// TwinCAT 3 PLC project KFEArbiter
// Title: KFE-ARBITER
// Company: SLAC - LCLS
// ProjectVersion: 0.0.0
// ProgramVersion: 3.1.4022.7
// CompilerDefines: K
// libraries:
//   PMPS, * (SLAC - LCLS)
//   Tc2_Math, * (Beckhoff Automation GmbH)
//   Tc2_MC2, * (Beckhoff Automation GmbH)
//   Tc2_Standard, * (Beckhoff Automation GmbH)
//   Tc2_System, * (Beckhoff Automation GmbH)
//   Tc2_SystemCX, * (Beckhoff Automation GmbH)
//   Tc2_Utilities, * (Beckhoff Automation GmbH)
//   Tc3_Module, * (Beckhoff Automation GmbH)
//   LCLS General,2.8.2,SLAC
// project tree:
//   / FFOTask.TcTTO, PlcTask.TcTTO
//   GVLs/ GVL.TcGVL, GVL_CheckBounds.TcGVL
//   ImplicitChecks/ CheckBounds.TcPOU, CheckRangeSigned.TcPOU, CheckRangeUnsigned.TcPOU
//   POUs/ CurrentBPUpdate.TcPOU, CXDisplay.TcPOU, Fast_Faults_Evaluate.TcPOU, FB_BeamClassOutputs.TcPOU, MachineSimulation.TcPOU, MAIN.TcPOU, PMPS_Arbiter.TcPOU, P_AT1K0_SL1K0.TcPOU, P_BeamClassAssertion.TcPOU, P_Override_Tran_BC.TcPOU, P_SATT.TcPOU, Testing.TcPOU
//   POUs/TEMP/ FB_ArbiterToSubSys_IO.TcPOU
// real-time tasks:
//   TASK PlcTask: cycle T#10ms, priority 2, ADS port 350
//   TASK FFOTask: cycle T#1ms, priority 1, ADS port 351
// I/O:
//   DEVICE Device 1 (EtherCAT), AmsNetId 0.0.0.0.2.1
//     E0 (EK1200) [EK1200-5000 EtherCAT Power supply (2A E-Bus)]
//       FFO [EL2202 2Ch. Dig. Output 24V, 0.5A]
//       PMPS_Premp [EL2809 16Ch. Dig. Output 24V, 0.5A]
//       E3 (EK1122) [EK1122 2 port EtherCAT junction]
//         950-101W-R4-MPS-2 [EK1100 EtherCAT Coupler (2A E-Bus)]
//           PPS Stoppers 1 [EL1008 8Ch. Dig. Input 24V, 3ms]
//           PPS Stoppers 2 [EL1008 8Ch. Dig. Input 24V, 3ms]
//           950-101W-R4-MPS-2-E3 (EL9011) [EL9011 End Terminal]
//       Term 22 (EK1110) [EK1110 EtherCAT extension]
//     B940-009-R07-MPS-1 CU1-ESC1 [CU1128 6x EtherCAT junction]
//       plc-kfe-motion [EL6695 EtherCAT Bridge terminal (Secondary)]
//       plc-kfe-gmd-vac-01 [EL6695 EtherCAT Bridge terminal (Secondary)]
//       plc-kfe-xgmd-vac-01 [EL6695 EtherCAT Bridge terminal (Secondary)]
//       plc-kfe-vac [EL6692 EtherCAT Bridge terminal (Secondary)]
//       plc-kfe-gatt [EL6695 EtherCAT Bridge terminal (Secondary)]
//       plc-tmo-mot [EL6692 EtherCAT Bridge terminal (Secondary)]
//       plc-tmo-optics [EL6695 EtherCAT Bridge terminal (Secondary)]
//       plc-tmo-vac [EL6692 EtherCAT Bridge terminal (Secondary)]
//       B940-009-R07-MPS-1 CU1-ESC2 [CU1128 6x EtherCAT junction - Dev A]
//         plc-rix-mot
//         plc-rix-vac
//         plc-rix-optics
//         plc-crix-vac
//         plc-crix-mot
//       B940-009-R07-MPS-1 CU1-ESC3 [CU1128 6x EtherCAT junction - Dev B]
//         plc-qrix-vac
//         plc-qrix-mot
//         plc-txi-optics
//     plc-txi-mot [EL6695 EtherCAT Bridge terminal (Secondary)]
//     plc-txi-vac [EL6695 EtherCAT Bridge terminal (Secondary)]
// variable links:
//   KFEArbiter Instance <-> Device 1 (EtherCAT)
//     PlcTask Inputs/MAIN.fbEcatDiag.arrEcMasterNetId <-> InfoData/AmsNetId
//     PlcTask Inputs/MAIN.fbEcatDiag.nEcMasterDevState <-> Inputs/DevState
//     PlcTask Inputs/MAIN.fbEcatDiag.nEcMasterDeviceId <-> InfoData/DevId
//     PlcTask Inputs/MAIN.fbEcatDiag.nEcMasterSlaveCount <-> Inputs/SlaveCount
//     PlcTask Inputs/MAIN.fbEcatDiag.nEcMasterSlaveCountCfg <-> InfoData/CfgSlaveCount
//     PlcTask Inputs/MAIN.fbEcatDiag.wFrmXWcState <-> Inputs/Frm1WcState
//   KFEArbiter Instance <-> Device 1 (EtherCAT)/B940-009-R07-MPS-1 CU1-ESC1/B940-009-R07-MPS-1 CU1-ESC2/plc-crix-mot
//     PlcTask Inputs/PMPS_Arbiter.plc_crix_mot_PMPS_IO.i_Connected <-> SYNC Inputs/External device not connected
//     PlcTask Inputs/PMPS_Arbiter.plc_crix_mot_PMPS_IO.i_RequestedBP <-> IO Inputs/RequestedBP
//     PlcTask Inputs/PMPS_Arbiter.plc_crix_mot_PMPS_IO.i_TxPDOState <-> SYNC Inputs/TxPDO state
//     PlcTask Inputs/PMPS_Arbiter.plc_crix_mot_PMPS_IO.i_WcState <-> WcState/WcStateIn
//     PlcTask Outputs/PMPS_Arbiter.plc_crix_mot_PMPS_IO.o_CurrentBP <-> IO Outputs/CurrentBP
//   KFEArbiter Instance <-> Device 1 (EtherCAT)/B940-009-R07-MPS-1 CU1-ESC1/B940-009-R07-MPS-1 CU1-ESC2/plc-crix-vac
//     PlcTask Inputs/PMPS_Arbiter.plc_crix_vac_PMPS_IO.i_Connected <-> SYNC Inputs/External device not connected
//     PlcTask Inputs/PMPS_Arbiter.plc_crix_vac_PMPS_IO.i_RequestedBP <-> IO Inputs/RequestedBP
//     PlcTask Inputs/PMPS_Arbiter.plc_crix_vac_PMPS_IO.i_TxPDOState <-> SYNC Inputs/TxPDO state
//     PlcTask Inputs/PMPS_Arbiter.plc_crix_vac_PMPS_IO.i_WcState <-> WcState/WcStateIn
//     PlcTask Outputs/PMPS_Arbiter.plc_crix_vac_PMPS_IO.o_CurrentBP <-> IO Outputs/CurrentBP
//   KFEArbiter Instance <-> Device 1 (EtherCAT)/B940-009-R07-MPS-1 CU1-ESC1/B940-009-R07-MPS-1 CU1-ESC2/plc-rix-mot
//     PlcTask Inputs/PMPS_Arbiter.plc_rix_mot_PMPS_IO.i_Connected <-> SYNC Inputs/External device not connected
//     PlcTask Inputs/PMPS_Arbiter.plc_rix_mot_PMPS_IO.i_RequestedBP <-> IO Inputs/RequestedBP
//     PlcTask Inputs/PMPS_Arbiter.plc_rix_mot_PMPS_IO.i_TxPDOState <-> SYNC Inputs/TxPDO state
//     PlcTask Inputs/PMPS_Arbiter.plc_rix_mot_PMPS_IO.i_WcState <-> WcState/WcStateIn
//     PlcTask Inputs/P_SATT.i_SattArrayStatus_RIX <-> IO Inputs/SattArrayStatus
//     PlcTask Inputs/P_SATT.i_bWcStateIn_rix_mot <-> WcState/WcStateIn
//     PlcTask Inputs/P_SATT.i_bWcStateOut_rix_mot <-> WcState/WcStateOut
//     PlcTask Inputs/P_SATT.i_nState_rix_mot <-> InfoData/State
//     PlcTask Outputs/PMPS_Arbiter.plc_rix_mot_PMPS_IO.o_CurrentBP <-> IO Outputs/CurrentBP
//     PlcTask Outputs/P_SATT.q_SattArrayReq <-> IO Outputs/SattArrayReq
//   KFEArbiter Instance <-> Device 1 (EtherCAT)/B940-009-R07-MPS-1 CU1-ESC1/B940-009-R07-MPS-1 CU1-ESC2/plc-rix-optics
//     PlcTask Inputs/CurrentBPUpdate.i_MR1K1_ENC <-> IO Inputs/MR1K1_Y_ENC
//     PlcTask Inputs/PMPS_Arbiter.plc_rix_optics_PMPS_IO.i_Connected <-> SYNC Inputs/External device not connected
//     PlcTask Inputs/PMPS_Arbiter.plc_rix_optics_PMPS_IO.i_RequestedBP <-> IO Inputs/RequestedBP
//     PlcTask Inputs/PMPS_Arbiter.plc_rix_optics_PMPS_IO.i_TxPDOState <-> SYNC Inputs/TxPDO state
//     PlcTask Inputs/PMPS_Arbiter.plc_rix_optics_PMPS_IO.i_WcState <-> WcState/WcStateIn
//     PlcTask Outputs/PMPS_Arbiter.plc_rix_optics_PMPS_IO.o_CurrentBP <-> IO Outputs/CurrentBP
//   KFEArbiter Instance <-> Device 1 (EtherCAT)/B940-009-R07-MPS-1 CU1-ESC1/B940-009-R07-MPS-1 CU1-ESC2/plc-rix-vac
//     PlcTask Inputs/PMPS_Arbiter.plc_rix_vac_PMPS_IO.i_Connected <-> SYNC Inputs/External device not connected
//     PlcTask Inputs/PMPS_Arbiter.plc_rix_vac_PMPS_IO.i_RequestedBP <-> IO Inputs/RequestedBP
//     PlcTask Inputs/PMPS_Arbiter.plc_rix_vac_PMPS_IO.i_TxPDOState <-> SYNC Inputs/TxPDO state
//     PlcTask Inputs/PMPS_Arbiter.plc_rix_vac_PMPS_IO.i_WcState <-> WcState/WcStateIn
//     PlcTask Outputs/PMPS_Arbiter.plc_rix_vac_PMPS_IO.o_CurrentBP <-> IO Outputs/CurrentBP
//   KFEArbiter Instance <-> Device 1 (EtherCAT)/B940-009-R07-MPS-1 CU1-ESC1/B940-009-R07-MPS-1 CU1-ESC3/plc-qrix-mot
//     PlcTask Inputs/PMPS_Arbiter.plc_qrix_mot_PMPS_IO.i_Connected <-> SYNC Inputs/External device not connected
//     PlcTask Inputs/PMPS_Arbiter.plc_qrix_mot_PMPS_IO.i_RequestedBP <-> IO Inputs/RequestedBP
//     PlcTask Inputs/PMPS_Arbiter.plc_qrix_mot_PMPS_IO.i_TxPDOState <-> SYNC Inputs/TxPDO state
//     PlcTask Inputs/PMPS_Arbiter.plc_qrix_mot_PMPS_IO.i_WcState <-> WcState/WcStateIn
//     PlcTask Outputs/PMPS_Arbiter.plc_qrix_mot_PMPS_IO.o_CurrentBP <-> IO Outputs/CurrentBP
//   KFEArbiter Instance <-> Device 1 (EtherCAT)/B940-009-R07-MPS-1 CU1-ESC1/B940-009-R07-MPS-1 CU1-ESC3/plc-qrix-vac
//     PlcTask Inputs/Fast_Faults_Evaluate.i_xFastFaultOut_qrix_vac <-> IO Inputs/FFO
//     PlcTask Inputs/PMPS_Arbiter.plc_qrix_vac_PMPS_IO.i_Connected <-> SYNC Inputs/External device not connected
//     PlcTask Inputs/PMPS_Arbiter.plc_qrix_vac_PMPS_IO.i_RequestedBP <-> IO Inputs/RequestedBP
//     PlcTask Inputs/PMPS_Arbiter.plc_qrix_vac_PMPS_IO.i_TxPDOState <-> SYNC Inputs/TxPDO state
//     PlcTask Inputs/PMPS_Arbiter.plc_qrix_vac_PMPS_IO.i_WcState <-> WcState/WcStateIn
//     PlcTask Outputs/PMPS_Arbiter.plc_qrix_vac_PMPS_IO.o_CurrentBP <-> IO Outputs/CurrentBP
//   KFEArbiter Instance <-> Device 1 (EtherCAT)/B940-009-R07-MPS-1 CU1-ESC1/B940-009-R07-MPS-1 CU1-ESC3/plc-txi-optics
//     PlcTask Inputs/CurrentBPUpdate.i_MR1K3_ENC <-> IO Inputs/MR1K3_Y_ENC
//     PlcTask Inputs/CurrentBPUpdate.i_MR2K3_ENC <-> IO Inputs/MR2K3_Y_ENC
//     PlcTask Inputs/Fast_Faults_Evaluate.i_xFastFaultOut_txi_optics <-> IO Inputs/FFO
//     PlcTask Inputs/PMPS_Arbiter.plc_txi_optics_PMPS_IO.i_Connected <-> SYNC Inputs/External device not connected
//     PlcTask Inputs/PMPS_Arbiter.plc_txi_optics_PMPS_IO.i_RequestedBP <-> IO Inputs/RequestedBP
//     PlcTask Inputs/PMPS_Arbiter.plc_txi_optics_PMPS_IO.i_TxPDOState <-> SYNC Inputs/TxPDO state
//     PlcTask Inputs/PMPS_Arbiter.plc_txi_optics_PMPS_IO.i_WcState <-> WcState/WcStateIn
//     PlcTask Outputs/PMPS_Arbiter.plc_txi_optics_PMPS_IO.o_CurrentBP <-> IO Outputs/CurrentBP
//   KFEArbiter Instance <-> Device 1 (EtherCAT)/B940-009-R07-MPS-1 CU1-ESC1/plc-kfe-gatt
//     PlcTask Inputs/PMPS_Arbiter.plc_kfe_gatt_PMPS_IO.i_Connected <-> SYNC Inputs/External device not connected
//     PlcTask Inputs/PMPS_Arbiter.plc_kfe_gatt_PMPS_IO.i_RequestedBP <-> IO Inputs/RequestedBP
//     PlcTask Inputs/PMPS_Arbiter.plc_kfe_gatt_PMPS_IO.i_TxPDOState <-> SYNC Inputs/TxPDO state
//     PlcTask Inputs/PMPS_Arbiter.plc_kfe_gatt_PMPS_IO.i_WcState <-> WcState/WcStateIn
//     PlcTask Inputs/P_AT1K0_SL1K0.i_bWcStateIn_AT1K0 <-> WcState/WcStateIn
//     PlcTask Inputs/P_AT1K0_SL1K0.i_bWcStateOut_AT1K0 <-> WcState/WcStateOut
//     PlcTask Inputs/P_AT1K0_SL1K0.i_nState_AT1K0 <-> InfoData/State
//     PlcTask Inputs/P_AT1K0_SL1K0.i_nTranToAT1K0Stat <-> IO Inputs/Current Transmission
//     PlcTask Outputs/PMPS_Arbiter.plc_kfe_gatt_PMPS_IO.o_CurrentBP <-> IO Outputs/CurrentBP
//     PlcTask Outputs/P_AT1K0_SL1K0.q_nTranToAT1K0Req <-> IO Outputs/Requested Transmission
//   KFEArbiter Instance <-> Device 1 (EtherCAT)/B940-009-R07-MPS-1 CU1-ESC1/plc-kfe-gmd-vac-01
//     PlcTask Inputs/PMPS_Arbiter.plc_kfe_gmd_PMPS_IO.i_Connected <-> SYNC Inputs/External device not connected
//     PlcTask Inputs/PMPS_Arbiter.plc_kfe_gmd_PMPS_IO.i_RequestedBP <-> IO Inputs/RequestedBP
//     PlcTask Inputs/PMPS_Arbiter.plc_kfe_gmd_PMPS_IO.i_TxPDOState <-> SYNC Inputs/TxPDO state
//     PlcTask Inputs/PMPS_Arbiter.plc_kfe_gmd_PMPS_IO.i_WcState <-> WcState/WcStateIn
//     PlcTask Outputs/PMPS_Arbiter.plc_kfe_gmd_PMPS_IO.o_CurrentBP <-> IO Outputs/CurrentBP
//   KFEArbiter Instance <-> Device 1 (EtherCAT)/B940-009-R07-MPS-1 CU1-ESC1/plc-kfe-motion
//     PlcTask Inputs/CurrentBPUpdate.ST1K4_Y_ENC <-> IO Inputs/ST1K4_Y_ENC
//     PlcTask Inputs/PMPS_Arbiter.plc_kfe_motion_PMPS_IO.i_Connected <-> SYNC Inputs/External device not connected
//     PlcTask Inputs/PMPS_Arbiter.plc_kfe_motion_PMPS_IO.i_RequestedBP <-> IO Inputs/RequestedBP
//     PlcTask Inputs/PMPS_Arbiter.plc_kfe_motion_PMPS_IO.i_TxPDOState <-> SYNC Inputs/TxPDO state
//     PlcTask Inputs/PMPS_Arbiter.plc_kfe_motion_PMPS_IO.i_WcState <-> WcState/WcStateIn
//     PlcTask Inputs/P_AT1K0_SL1K0.i_bWcStateIn_KFEMOT <-> WcState/WcStateIn
//     PlcTask Inputs/P_AT1K0_SL1K0.i_bWcStateOut_KFEMOT <-> WcState/WcStateOut
//     PlcTask Inputs/P_AT1K0_SL1K0.i_nState_KFEMOT <-> InfoData/State
//     PlcTask Inputs/P_AT1K0_SL1K0.i_stAptArrayStat <-> IO Inputs/AptArrayStatus
//     PlcTask Inputs/P_SATT.i_SattArrayStatus_KFE <-> IO Inputs/SattArrayStatus
//     PlcTask Inputs/P_SATT.i_bWcStateIn_kfe_mot <-> WcState/WcStateIn
//     PlcTask Inputs/P_SATT.i_bWcStateOut_kfe_mot <-> WcState/WcStateOut
//     PlcTask Inputs/P_SATT.i_nState_kfe_mot <-> InfoData/State
//     PlcTask Outputs/PMPS_Arbiter.plc_kfe_motion_PMPS_IO.o_CurrentBP <-> IO Outputs/CurrentBP
//     PlcTask Outputs/P_AT1K0_SL1K0.q_stAptArrayReq <-> IO Outputs/AptArrayReq
//   KFEArbiter Instance <-> Device 1 (EtherCAT)/B940-009-R07-MPS-1 CU1-ESC1/plc-kfe-vac
//     PlcTask Inputs/PMPS_Arbiter.plc_kfe_vac_PMPS_IO.i_Connected <-> SYNC Inputs/External device not connected
//     PlcTask Inputs/PMPS_Arbiter.plc_kfe_vac_PMPS_IO.i_RequestedBP <-> IO Inputs/RequestedBP
//     PlcTask Inputs/PMPS_Arbiter.plc_kfe_vac_PMPS_IO.i_TxPDOState <-> SYNC Inputs/TxPDO state
//     PlcTask Inputs/PMPS_Arbiter.plc_kfe_vac_PMPS_IO.i_WcState <-> WcState/WcStateIn
//     PlcTask Outputs/PMPS_Arbiter.plc_kfe_vac_PMPS_IO.o_CurrentBP <-> IO Outputs/CurrentBP
//   KFEArbiter Instance <-> Device 1 (EtherCAT)/B940-009-R07-MPS-1 CU1-ESC1/plc-kfe-xgmd-vac-01
//     PlcTask Inputs/PMPS_Arbiter.plc_kfe_xgmd_PMPS_IO.i_Connected <-> SYNC Inputs/External device not connected
//     PlcTask Inputs/PMPS_Arbiter.plc_kfe_xgmd_PMPS_IO.i_RequestedBP <-> IO Inputs/RequestedBP
//     PlcTask Inputs/PMPS_Arbiter.plc_kfe_xgmd_PMPS_IO.i_TxPDOState <-> SYNC Inputs/TxPDO state
//     PlcTask Inputs/PMPS_Arbiter.plc_kfe_xgmd_PMPS_IO.i_WcState <-> WcState/WcStateIn
//     PlcTask Outputs/PMPS_Arbiter.plc_kfe_xgmd_PMPS_IO.o_CurrentBP <-> IO Outputs/CurrentBP
//   KFEArbiter Instance <-> Device 1 (EtherCAT)/B940-009-R07-MPS-1 CU1-ESC1/plc-tmo-mot
//     PlcTask Inputs/CurrentBPUpdate.st4k4Watcher.i_StopperInLS <-> IO Inputs/bST4K4_IN
//     PlcTask Inputs/CurrentBPUpdate.st4k4Watcher.i_StopperOutLS <-> IO Inputs/bST4K4_OUT
//     PlcTask Inputs/PMPS_Arbiter.plc_tmo_motion_PMPS_IO.i_Connected <-> SYNC Inputs/External device not connected
//     PlcTask Inputs/PMPS_Arbiter.plc_tmo_motion_PMPS_IO.i_RequestedBP <-> IO Inputs/RequestedBP
//     PlcTask Inputs/PMPS_Arbiter.plc_tmo_motion_PMPS_IO.i_TxPDOState <-> SYNC Inputs/TxPDO state
//     PlcTask Inputs/PMPS_Arbiter.plc_tmo_motion_PMPS_IO.i_WcState <-> WcState/WcStateIn
//     PlcTask Outputs/PMPS_Arbiter.plc_tmo_motion_PMPS_IO.o_CurrentBP <-> IO Outputs/CurrentBP
//   KFEArbiter Instance <-> Device 1 (EtherCAT)/B940-009-R07-MPS-1 CU1-ESC1/plc-tmo-optics
//     PlcTask Inputs/PMPS_Arbiter.plc_tmo_optics_PMPS_IO.i_Connected <-> SYNC Inputs/External device not connected
//     PlcTask Inputs/PMPS_Arbiter.plc_tmo_optics_PMPS_IO.i_RequestedBP <-> IO Inputs/RequestedBP
//     PlcTask Inputs/PMPS_Arbiter.plc_tmo_optics_PMPS_IO.i_TxPDOState <-> SYNC Inputs/TxPDO state
//     PlcTask Inputs/PMPS_Arbiter.plc_tmo_optics_PMPS_IO.i_WcState <-> WcState/WcStateIn
//     PlcTask Outputs/PMPS_Arbiter.plc_tmo_optics_PMPS_IO.o_CurrentBP <-> IO Outputs/CurrentBP
//   KFEArbiter Instance <-> Device 1 (EtherCAT)/B940-009-R07-MPS-1 CU1-ESC1/plc-tmo-vac
//     PlcTask Inputs/PMPS_Arbiter.plc_tmo_vacuum_PMPS_IO.i_Connected <-> SYNC Inputs/External device not connected
//     PlcTask Inputs/PMPS_Arbiter.plc_tmo_vacuum_PMPS_IO.i_RequestedBP <-> IO Inputs/RequestedBP
//     PlcTask Inputs/PMPS_Arbiter.plc_tmo_vacuum_PMPS_IO.i_TxPDOState <-> SYNC Inputs/TxPDO state
//     PlcTask Inputs/PMPS_Arbiter.plc_tmo_vacuum_PMPS_IO.i_WcState <-> WcState/WcStateIn
//     PlcTask Outputs/PMPS_Arbiter.plc_tmo_vacuum_PMPS_IO.o_CurrentBP <-> IO Outputs/CurrentBP
//   KFEArbiter Instance <-> Device 1 (EtherCAT)/E0 (EK1200)/E3 (EK1122)/950-101W-R4-MPS-2/PPS Stoppers 1
//     PlcTask Inputs/CurrentBPUpdate.st1k2Watcher.i_StopperInLS <-> Channel 3/ST1K2 IN
//     PlcTask Inputs/CurrentBPUpdate.st1k3Watcher.i_StopperInLS <-> Channel 5/ST1K3 IN
//     PlcTask Inputs/CurrentBPUpdate.st3k4Watcher.i_StopperInLS <-> Channel 1/ST3K4 IN
//     PlcTask Inputs/CurrentBPUpdate.st1k2Watcher.i_StopperOutLS <-> Channel 4/ST1K2 OUT
//     PlcTask Inputs/CurrentBPUpdate.st1k3Watcher.i_StopperOutLS <-> Channel 6/ST1K3 OUT
//     PlcTask Inputs/CurrentBPUpdate.st3k4Watcher.i_StopperOutLS <-> Channel 2/ST3K4 OUT
//   KFEArbiter Instance <-> Device 1 (EtherCAT)/E0 (EK1200)/FFO
//     PlcTask Outputs/GVL.g_FastFaultOutput1.q_xFastFaultOut <-> Channel 1/Output
//     PlcTask Outputs/GVL.g_FastFaultOutput2.q_xFastFaultOut <-> Channel 2/Output
//   KFEArbiter Instance <-> Device 1 (EtherCAT)/E0 (EK1200)/PMPS_Premp
//     PlcTask Outputs/CurrentBPUpdate.q_MR1K1_VETO <-> Channel 13/MR1K1 IN
//     PlcTask Outputs/CurrentBPUpdate.st1k2Watcher.q_StopperIN_Relay <-> Channel 14/ST1K2 RELAY IN
//     PlcTask Outputs/CurrentBPUpdate.st1k3Watcher.q_StopperIN_Relay <-> Channel 7/ST1K3 RELAY IN
//     PlcTask Outputs/CurrentBPUpdate.st3k4Watcher.q_StopperIN_Relay <-> Channel 12/ST3K4 RELAY IN
//     PlcTask Outputs/MAIN.bM1K1_OUT_Override <-> Channel 8/Output
//     PlcTask Outputs/PMPS_Arbiter.fbCuInterface.q_CLTS_ASSERTION_LINES[1] <-> Channel 9/Output
//     PlcTask Outputs/PMPS_Arbiter.fbCuInterface.q_CLTS_ASSERTION_LINES[2] <-> Channel 10/Output
//     PlcTask Outputs/PMPS_Arbiter.fbCuInterface.q_CLTS_ASSERTION_LINES[3] <-> Channel 11/Output
//     PlcTask Outputs/P_BeamClassAssertion.fbMPSInterface.q_BC_ASSERTION_LINES[{1..4}] <-> Channel {1..4}/Output  (4 links)
//   KFEArbiter Instance <-> Device 1 (EtherCAT)/plc-txi-mot
//     PlcTask Inputs/Fast_Faults_Evaluate.i_xFastFaultOut_txi_mot <-> IO Inputs/FFO
//     PlcTask Inputs/PMPS_Arbiter.plc_txi_motion_PMPS_IO.i_Connected <-> SYNC Inputs/External device not connected
//     PlcTask Inputs/PMPS_Arbiter.plc_txi_motion_PMPS_IO.i_RequestedBP <-> IO Inputs/RequestedBP
//     PlcTask Inputs/PMPS_Arbiter.plc_txi_motion_PMPS_IO.i_TxPDOState <-> SYNC Inputs/TxPDO state
//     PlcTask Inputs/PMPS_Arbiter.plc_txi_motion_PMPS_IO.i_WcState <-> WcState/WcStateIn
//     PlcTask Outputs/PMPS_Arbiter.plc_txi_motion_PMPS_IO.o_CurrentBP <-> IO Outputs/CurrentBP
//   KFEArbiter Instance <-> Device 1 (EtherCAT)/plc-txi-vac
//     PlcTask Inputs/Fast_Faults_Evaluate.i_xFastFaultOut_txi_vac <-> IO Inputs/FFO
//     PlcTask Inputs/PMPS_Arbiter.plc_txi_vacuum_PMPS_IO.i_Connected <-> SYNC Inputs/External device not connected
//     PlcTask Inputs/PMPS_Arbiter.plc_txi_vacuum_PMPS_IO.i_RequestedBP <-> IO Inputs/RequestedBP
//     PlcTask Inputs/PMPS_Arbiter.plc_txi_vacuum_PMPS_IO.i_TxPDOState <-> SYNC Inputs/TxPDO state
//     PlcTask Inputs/PMPS_Arbiter.plc_txi_vacuum_PMPS_IO.i_WcState <-> WcState/WcStateIn
//     PlcTask Outputs/PMPS_Arbiter.plc_txi_vacuum_PMPS_IO.o_CurrentBP <-> IO Outputs/CurrentBP

CONFIGURATION KFEArbiter
    RESOURCE PLC ON TwinCAT3
        TASK FFOTask(INTERVAL := T#1ms, PRIORITY := 1);
        TASK PlcTask(INTERVAL := T#10ms, PRIORITY := 2);
        PROGRAM MAIN WITH PlcTask : MAIN;
    END_RESOURCE
END_CONFIGURATION

// ---- GVLs/GVL.TcGVL

VAR_GLOBAL
   {attribute 'pytmc' := '
    pv: @(PREFIX)Arbiter:01
    '}
    g_fbArbiter1	:	FB_Arbiter(25);

    {attribute 'pytmc' := '
    pv: @(PREFIX)Arbiter:02
    '}
    g_fbArbiter2	:	FB_Arbiter(25); //Used to line beam parameter

    ReqBP	:	ST_BeamParams; //Currently the placeholder for the fully arbitrated BP set

    // These are added for the additional low selector to figure out the override
    stArbiter1BP:ST_BeamParams; // a place holder for the arbitrated safe beam set from all the connected PLCs
    stCurrentFakeBP:ST_BeamParams; //Currently the placeholder for the fake arbitrated BP set to go to the rest of the PLC

    {attribute 'pytmc' := '
    pv: @(PREFIX)FFO:01
    '}
    {attribute 'TcLinkTo' := '.q_xFastFaultOut:=TIIB[FFO]^Channel 1^Output'}
    g_FastFaultOutput1	:	FB_HardwareFFOutput := (bAutoReset:=TRUE);

    {attribute 'pytmc' := '
    pv: @(PREFIX)FFO:02
    '}
    {attribute 'TcLinkTo' := '.q_xFastFaultOut:=TIIB[FFO]^Channel 2^Output'}
    g_FastFaultOutput2	:	FB_HardwareFFOutput := (bAutoReset:=TRUE);
	
	
	//The following faults will be per hutch and vetoed by the hutch specific veto
	//TMO OPTICS, VAC and Motion, DREAM
	{attribute 'pytmc' := '
    pv: @(PREFIX)FFO:03
    '}
    g_FastFaultOutput3	:	FB_HardwareFFOutput := (bAutoReset:=TRUE);
	{attribute 'pytmc' := '
    pv: @(PREFIX)FFO:04
    '}
    g_FastFaultOutput4	:	FB_HardwareFFOutput := (bAutoReset:=TRUE);
	
	
	//RIX Motion, QRIX and CRIX
	//NOTE: NOT OPTICS, NO VETO for OPTICS
	{attribute 'pytmc' := '
    pv: @(PREFIX)FFO:05
    '}
    g_FastFaultOutput5	:	FB_HardwareFFOutput := (bAutoReset:=TRUE);
	
	{attribute 'pytmc' := '
    pv: @(PREFIX)FFO:06
    '}
    g_FastFaultOutput6	:	FB_HardwareFFOutput := (bAutoReset:=TRUE);
	
	
	//TXI VAC and MOTION 
	//NOTE: NOT OPTICS, NO VETO for OPTICS
	{attribute 'pytmc' := '
    pv: @(PREFIX)FFO:07
    '}
    g_FastFaultOutput7	:	FB_HardwareFFOutput := (bAutoReset:=TRUE);
	

    g_rTestingVelocity	:	LREAL := PMPS_GVL.VISIBLE_TEST_VELOCITY;

     {attribute 'pytmc' := '
       pv: @(PREFIX)ApplyJF
    '}
    bApplyJF: BOOL:=FALSE;
    // Administrative mode for beam intensity
     {attribute 'pytmc' := '
          pv: @(PREFIX)IntensityJF
    '}
    nBeamIntensityJF: REAL :=nBeamIntensity;

    {attribute 'pytmc' := '
          pv: @(PREFIX)CancelJF
    '}
    bCancelJF: BOOL:=FALSE;

    {attribute 'pytmc' := '
          pv: @(PREFIX)DurationJF
    '}
    rDurationJF: REAL:=GVL.MaxDuration;//hours

    {attribute 'pytmc' := '
          pv: @(PREFIX)TimeRemainJF
    '}
    rTimeRemainJF: REAL:=GVL.MaxDuration;//hours

    AttemptReset    :   BOOL; // For testing
END_VAR

VAR_GLOBAL CONSTANT
    MAX_FAST_FAULTS : UINT := 100;
    //Judgement factor constants (administrative mode)
    nBeamIntensity : INT :=5;//mj
    MaxDuration : REAL :=12;

END_VAR

// ---- GVLs/GVL_CheckBounds.TcGVL
{attribute 'qualified_only'}
VAR_GLOBAL
    nTooLow : UDINT;
    nTooHigh : UDINT;
    nDivByZero : UDINT;
END_VAR

// ---- POUs/MAIN.TcPOU
PROGRAM MAIN
VAR
    Initialize	:	BOOL := TRUE;

    fbLogHandler : FB_LogHandler;
    fbEcatDiag : FB_EcatDiagWrapper;



    PERanges : PE_Ranges;
    {attribute 'TcLinkTo' := 'TIIB[PMPS_Premp]^Channel 8^Output;'}
    bM1K1_OUT_Override AT %Q* : BOOL; // Using this book to completely overrule the last bit of the BC interface.

    //System Time
     {attribute 'pytmc' := '
        pv: @(PREFIX)SystemDT
        io: i
     '}
    SystemTime:DINT;
    fbTime : FB_LocalSystemTime := ( bEnable := TRUE, dwCycle := 1 ); //Get current system time, used for override
    fbTime_to_UTC: FB_TzSpecificLocalTimeToSystemTime;
    fbGetTimeZone: FB_GetTimeZoneInformation;
END_VAR

//Arbiter PLC

IF Initialize THEN
    Initialize := FALSE;
END_IF

// Ethercat Diagnostics
fbEcatDiag();

// PMPS Functionality
CurrentBPUpdate();

///////////////////////////////////////////////////
// This code should be disabled or removed in deployment
// Might have a switch to change to simulation mode
MachineSimulation();
//Testing();
///////////////////////////////////////////////////

PMPS_Arbiter();

P_AT1K0_SL1K0();

P_SATT();


bM1K1_OUT_Override := PMPS_GVL.stCurrentBeamParameters.aVetoDevices[PMPS.K_Stopper.MR1K1_OUT];

fbLogHandler();
A_SystemTime();
Fast_Faults_Evaluate();

ACTION A_SystemTime:
//Get local System Time
fbTime(sNetID:='');
//Get Time Zone
fbGetTimeZone(sNetID:='',bExecute:=TRUE,tTimeout:=T#10S);
//change local time to UTC to be compatible with unix time epoch widget
fbTime_to_UTC(in:= fbTime.systemTime , tzInfo:=fbGetTimeZone.tzInfo);

SystemTime:= TO_DINT(TO_DT(SystemTime_TO_DT(fbTime_to_UTC.out)));
END_ACTION

ACTION Initialize:

END_ACTION

END_PROGRAM

// ---- POUs/CurrentBPUpdate.TcPOU
PROGRAM CurrentBPUpdate
VAR
    {attribute 'pytmc' := '
        pv: @(PREFIX)K:Rate
        link: IOC:BSY0:MP01:BYKIKS_RATE
        field: EGU RateEnum
    '}
    fbBYKIK_Rate : FB_LREALFromEPICS := (
        iMaximumValidSeverity := 2);


    {attribute 'pytmc' := '
        pv: @(PREFIX)
    '}
    fbEPICS_KRate : FB_RateFromEPICS;

    {attribute 'pytmc' := '
        pv: @(PREFIX)L:BC
        link: SIOC:SYS0:MP03:SC_SXR_BC
        field: EGU BCEnum
    '}
    fbMPS_BeamClass : FB_LREALFromEPICS := (
        iMaximumValidSeverity := 2);

        {attribute 'pytmc' := '
        pv: @(PREFIX)
    '}
    fbEPICSKBeamClass : FB_BeamClassFromEPICS;

    {attribute 'pytmc' := '
        pv: @(PREFIX)K:Mode
        link: SIOC:FEES:MP01:FACMODE_RBV
    '}
    fbSXR_MachineMode : FB_LREALFromEPICS := (
        iMaximumValidSeverity := 2);

    {attribute 'pytmc' := '
        pv: @(PREFIX)
    '}
    fbEPICSLMachineMode : FB_MachineModeFromEPICS;

    {attribute 'pytmc' := '
        pv: @(PREFIX)PE
    '}
    fbKPhotonEnergy : FB_KPhotonEnergy;

    // Photon energy for the masses
    {attribute 'TcLinkTo' := 'TIIB[plc-kfe-gatt]^IO Outputs^rPhotonEnergy'}
    {attribute 'TcLinkTo' := 'TIIB[plc-rix-mot]^IO Outputs^rPhotonEnergy'}
    {attribute 'TcLinkTo' := 'TIIB[plc-rix-optics]^IO Outputs^rPhotonEnergy'}
    q_rPhotonEnergy AT %Q* : REAL;


    // Stoppers

    {attribute 'TcLinkTo' := '
                .i_StopperInLS:=TIIB[PPS Stoppers 1]^Channel 1^ST3K4 IN;
                .i_StopperOutLS:=TIIB[PPS Stoppers 1]^Channel 2^ST3K4 OUT;
                .q_StopperIN_Relay:=TIIB[PMPS_Premp]^Channel 12^ST3K4 RELAY IN;
                                '}
    st3k4Watcher : FB_KStopper(
        PMPS.K_Stopper.ST3K4,
        'ST3K4');

   {attribute 'TcLinkTo' := '
                .i_StopperInLS:=TIIB[PPS Stoppers 1]^Channel 3^ST1K2 IN;
                .i_StopperOutLS:=TIIB[PPS Stoppers 1]^Channel 4^ST1K2 OUT;
                .q_StopperIN_Relay:=TIIB[PMPS_Premp]^Channel 14^ST1K2 RELAY IN;
                                '}
    st1k2Watcher : FB_KStopper(
        PMPS.K_Stopper.ST1K2,
        'ST1K2');

    {attribute 'TcLinkTo' := '
                .i_StopperInLS:=TIIB[PPS Stoppers 1]^Channel 5^ST1K3 IN;
                .i_StopperOutLS:=TIIB[PPS Stoppers 1]^Channel 6^ST1K3 OUT;
                .q_StopperIN_Relay:=TIIB[PMPS_Premp]^Channel 7^ST1K3 RELAY IN;
                                '}
    st1k3Watcher : FB_KStopper(
        PMPS.K_Stopper.ST1K3,
        'ST1K3');

    // MR1K1 Veto
    ////////////////////////
          {attribute 'TcLinkTo' := 'TIIB[plc-rix-optics]^IO Inputs^MR1K1_Y_ENC'}
        i_MR1K1_ENC AT %I* : UDINT; // MR1K1 encoder from the rix optics system
        cMR1K1_IN_UpperLimit : UDINT := 33411000;
        cMR1K1_IN_LowerLimit : UDINT := 31911000;
        cMR1K1_OUT_UpperLimit : UDINT := 14173400;
        {attribute 'TcLinkTo' := 'TIIB[PMPS_Premp]^Channel 13^MR1K1 IN'}
        q_MR1K1_VETO AT %Q* : BOOL; // Signal to accel. MPS that MR1K1 is in
        fbMR1K1VetoDevice : FB_KVetoDevice(
            eVetoDeviceIN := K_Stopper.MR1K1_IN,
            eVetoDeviceOUT := K_Stopper.MR1K1_OUT,
            sVetoDeviceName := 'MR1K1');




    // ST4K4 Photon Terminator Veto
    {attribute 'TcLinkTo' := '
                .i_StopperInLS:=TIIB[plc-tmo-mot]^IO Inputs^bST4K4_IN;
                .i_StopperOutLS:=TIIB[plc-tmo-mot]^IO Inputs^bST4K4_OUT;
     '}
    st4k4Watcher : FB_KStopper(
        PMPS.K_Stopper.ST4K4,
        'ST4K4');


     // MR1K3 Veto
    ////////////////////////
          {attribute 'TcLinkTo' := 'TIIB[plc-txi-optics]^IO Inputs^MR1K3_Y_ENC'}
        i_MR1K3_ENC AT %I* : ULINT; // MR1K3 encoder from the txi k optics optics system
        cMR1K3_IN_UpperLimit : UDINT := 108500000 + 10000000;
        cMR1K3_IN_LowerLimit : UDINT := 108500000 - 10000000 ;
        cMR1K3_OUT_UpperLimit : UDINT := 8900000 + 100000;

        q_MR1K3_VETO AT %Q* : BOOL; // Signal to accel. MPS that MR1K3 is in
        fbMR1K3VetoDevice : FB_KVetoDevice(
            eVetoDeviceIN := K_Stopper.MR1K3_IN,
            eVetoDeviceOUT := K_Stopper.MR1K3_OUT,
            sVetoDeviceName := 'MR1K3');

    // MR2K3 Veto
    ////////////////////////
          {attribute 'TcLinkTo' := 'TIIB[plc-txi-optics]^IO Inputs^MR2K3_Y_ENC'}
        i_MR2K3_ENC AT %I* : ULINT; // MR2K3 encoder from the txi k optics system
        cMR2K3_IN_UpperLimit : UDINT := 105650000 + 10000000;
        cMR2K3_IN_LowerLimit : UDINT := 105650000 - 10000000 ;
        cMR2K3_OUT_UpperLimit : UDINT := 10000000;

        q_MR2K3_VETO AT %Q* : BOOL; // Signal to accel. MPS that MR2K3 is in
        fbMR2K3VetoDevice : FB_KVetoDevice(
            eVetoDeviceIN := K_Stopper.MR2K3_IN,
            eVetoDeviceOUT := K_Stopper.MR2K3_OUT,
            sVetoDeviceName := 'MR2K3');


    // ST1K4Veto
    // ST1K4 Test Photon stopper Veto in the FEE right before ST3K4 stopper
    st1k4Watcher :   FB_KVetoDevice(
            eVetoDeviceIN := K_Stopper.ST1K4,
            eVetoDeviceOUT := K_Stopper.DEFAULT, // not used there is no ST1K4 OUT Just a place holder
            sVetoDeviceName := 'ST1K4');
    ////////////////////////

          {attribute 'TcLinkTo' := 'TIIB[plc-kfe-motion]^IO Inputs^ST1K4_Y_ENC'}
        ST1K4_Y_ENC AT %I* : UDINT; // MR2K3 encoder from the  system
        ST1K4_IN_UpperLimit : UDINT := 4294002942 + 20000; //delta is 1mm
        ST1K4_IN_LowerLimit : UDINT := 4293982942;
        ST1K4_OUT_UpperLimit : UDINT := 8900000;

END_VAR

// Acquiring K-line rate
fbEPICS_KRate(BP:=PMPS_GVL.stCurrentBeamParameters, fbBYKIK_Rate:=fbBYKIK_Rate, FFO:=GVL.g_FastFaultOutput1);

// Acquiring photon energy
fbKPhotonEnergy(BP:=PMPS_GVL.stCurrentBeamParameters);

q_rPhotonEnergy := LREAL_TO_REAL(fbKPhotonEnergy.fbSXU.fCurrentPhotonEnergy);

//Update current photon energy
PMPS_GVL.stCurrentBeamParameters.neV := LREAL_TO_REAL(fbKPhotonEnergy.fbSXU.fCurrentPhotonEnergy);
// Acquiring K-line BeamClass
fbEPICSKBeamClass(BP:=PMPS_GVL.stCurrentBeamParameters, fbMPS_BeamClass:=fbMPS_BeamClass, FFO:=GVL.g_FastFaultOutput1);

// Acquiring K-line Machine Mode
fbEPICSLMachineMode(BP:=PMPS_GVL.stCurrentBeamParameters, fbMPS_MachineMode:=fbSXR_MachineMode, FFO:=GVL.g_FastFaultOutput1);


// Stopper readbacks
st3k4Watcher(stCurrentBP:=PMPS_GVL.stCurrentBeamParameters);
st1k2Watcher(stCurrentBP:=PMPS_GVL.stCurrentBeamParameters);
st1k3Watcher(stCurrentBP:=PMPS_GVL.stCurrentBeamParameters);
// ST4K4 Photon Terminator Veto
st4k4Watcher(stCurrentBP:=PMPS_GVL.stCurrentBeamParameters);
// MR1K1 Veto
////////////////////////
    fbMR1K1VetoDevice(
        i_bIn := cMR1K1_IN_LowerLimit < i_MR1K1_ENC	AND i_MR1K1_ENC < cMR1K1_IN_UpperLimit,
        i_bOut := i_MR1K1_ENC < cMR1K1_OUT_UpperLimit,
        q_bIN => q_MR1K1_VETO,
        stCurrentBP:= PMPS_GVL.stCurrentBeamParameters);

////////////////////////
    fbMR1K3VetoDevice(
        i_bIn := cMR1K3_IN_LowerLimit < i_MR1K3_ENC	AND i_MR1K3_ENC < cMR1K3_IN_UpperLimit,
        i_bOut := i_MR1K3_ENC < cMR1K3_OUT_UpperLimit,
        q_bIN => q_MR1K3_VETO,
        stCurrentBP:= PMPS_GVL.stCurrentBeamParameters);


// MR2K3 Veto
////////////////////////
    fbMR2K3VetoDevice(
        i_bIn := cMR2K3_IN_LowerLimit < i_MR2K3_ENC	AND i_MR2K3_ENC < cMR2K3_IN_UpperLimit,
        i_bOut := i_MR2K3_ENC < cMR2K3_OUT_UpperLimit,
        q_bIN => q_MR2K3_VETO,
        stCurrentBP:= PMPS_GVL.stCurrentBeamParameters);


// ST1K4 Photon Test stopper Veto
st1k4Watcher(i_bIn := ST1K4_IN_LowerLimit < ST1K4_Y_ENC	AND ST1K4_Y_ENC < ST1K4_IN_UpperLimit,
        i_bOut := ST1K4_Y_ENC <  ST1K4_OUT_UpperLimit,
        q_bIN => ,
        stCurrentBP:= PMPS_GVL.stCurrentBeamParameters);

END_PROGRAM

// ---- POUs/MachineSimulation.TcPOU
PROGRAM MachineSimulation
VAR
    fbMachine	:	FB_MachineSimulator; //Simulates attenuator as well
    fbeVSimulator : FB_eVSimulator := (NoiseLevel := 1);
END_VAR

// reV Simulator
fbeVSimulator();

// Machine simulator
fbMachine(
    i_stAssertedParams := PMPS_GVL.stRequestedBeamParameters,
    iq_stMachineParams := PMPS_GVL.stCurrentBeamParameters,
    i_xFault	:= NOT GVL.g_FastFaultOutput1.q_xFastFaultOut,
    xEnableAtt := false,
    xEnablePE := false
    );

//PMPS_GVL.stCurrentBeamParameters.neVRange := F_eVRangeCalculator(fbeVSimulator.eV, PMPS_GVL.stCurrentBeamParameters.neVRange);

//PMPS_GVL.stCurrentBeamParameters.neVRange := 0;

END_PROGRAM

// ---- POUs/PMPS_Arbiter.TcPOU
PROGRAM PMPS_Arbiter
VAR

    fbSetPE	:	PE_Ranges;

    fbBPRequestor : FB_BPRequestor; // Updates global PMPS RequestedBeamParams
    {attribute 'pytmc' := '
    pv: @(PREFIX)PhotonEnergyWatcher
    '}
    fbPhotonEnergyWatcher	:	FB_PhotonEnergyWatcher;

    {attribute 'pytmc' := '
    pv: @(PREFIX)CuRateOutputs
    '}
    fbCuInterface	:	FB_CTLS_Outputs;


    {attribute 'pytmc' := '
    pv: @(PREFIX)BeamParamCntl
    '}
    fbBPControl : FB_BPControlDevice(nID:=16#FFFF);

    (* Subsystem requests use this FB and a pragma link to pass their requests to the arbiter.
    The fb is called on each cycle and updates the arbiter with the current BP set requested
    from the subsystem PLC.*)
    //<TODO> make this so it does input and output to the IF
    (*{attribute 'pytmc' := '
    pv: @(PREFIX):PLC1
    '}*)
    {attribute 'TcLinkTo' := '.i_RequestedBP:=TIIB[plc-kfe-motion]^IO Inputs^RequestedBP;
                                .o_CurrentBP:=TIIB[plc-kfe-motion]^IO Outputs^CurrentBP;
                                .i_Connected:=TIIB[plc-kfe-motion]^SYNC Inputs^External device not connected;
                                .i_WcState:=TIIB[plc-kfe-motion]^WcState^WcStateIn;
                                .i_TxPDOState:=TIIB[plc-kfe-motion]^SYNC Inputs^TxPDO state;
                                '}
    plc_kfe_motion_PMPS_IO : FB_ArbiterToSubSys_IO := (RequestingSystemID := 16#FF0F);




    {attribute 'TcLinkTo' := '.i_RequestedBP:=TIIB[plc-kfe-vac]^IO Inputs^RequestedBP;
                                .o_CurrentBP:=TIIB[plc-kfe-vac]^IO Outputs^CurrentBP;
                                .i_Connected:=TIIB[plc-kfe-vac]^SYNC Inputs^External device not connected;
                                .i_WcState:=TIIB[plc-kfe-vac]^WcState^WcStateIn;
                                .i_TxPDOState:=TIIB[plc-kfe-vac]^SYNC Inputs^TxPDO state;
                                '}
    plc_kfe_vac_PMPS_IO : FB_ArbiterToSubSys_IO := (RequestingSystemID := 16#FF11);

    {attribute 'TcLinkTo' := '.i_RequestedBP:=TIIB[plc-kfe-gatt]^IO Inputs^RequestedBP;
                                .o_CurrentBP:=TIIB[plc-kfe-gatt]^IO Outputs^CurrentBP;
                                .i_Connected:=TIIB[plc-kfe-gatt]^SYNC Inputs^External device not connected;
                                .i_WcState:=TIIB[plc-kfe-gatt]^WcState^WcStateIn;
                                .i_TxPDOState:=TIIB[plc-kfe-gatt]^SYNC Inputs^TxPDO state;
                                '}
    plc_kfe_gatt_PMPS_IO : FB_ArbiterToSubSys_IO := (RequestingSystemID := 16#FF12);

    {attribute 'TcLinkTo' := '.i_RequestedBP:=TIIB[plc-kfe-gmd-vac-01]^IO Inputs^RequestedBP;
                                .o_CurrentBP:=TIIB[plc-kfe-gmd-vac-01]^IO Outputs^CurrentBP;
                                .i_Connected:=TIIB[plc-kfe-gmd-vac-01]^SYNC Inputs^External device not connected;
                                .i_WcState:=TIIB[plc-kfe-gmd-vac-01]^WcState^WcStateIn;
                                .i_TxPDOState:=TIIB[plc-kfe-gmd-vac-01]^SYNC Inputs^TxPDO state;
                                '}
    plc_kfe_gmd_PMPS_IO : FB_ArbiterToSubSys_IO := (RequestingSystemID := 16#FF13);

    {attribute 'TcLinkTo' := '.i_RequestedBP:=TIIB[plc-kfe-xgmd-vac-01]^IO Inputs^RequestedBP;
                                .o_CurrentBP:=TIIB[plc-kfe-xgmd-vac-01]^IO Outputs^CurrentBP;
                                .i_Connected:=TIIB[plc-kfe-xgmd-vac-01]^SYNC Inputs^External device not connected;
                                .i_WcState:=TIIB[plc-kfe-xgmd-vac-01]^WcState^WcStateIn;
                                .i_TxPDOState:=TIIB[plc-kfe-xgmd-vac-01]^SYNC Inputs^TxPDO state;
                                '}
    plc_kfe_xgmd_PMPS_IO : FB_ArbiterToSubSys_IO := (RequestingSystemID := 16#FF14);



//////////////////////////////////////////////
// TMO PLCs
/////////////////////////////////////////////

    {attribute 'TcLinkTo' := '.i_RequestedBP:=TIIB[plc-tmo-mot]^IO Inputs^RequestedBP;
                                .o_CurrentBP:=TIIB[plc-tmo-mot]^IO Outputs^CurrentBP;
                                .i_Connected:=TIIB[plc-tmo-mot]^SYNC Inputs^External device not connected;
                                .i_WcState:=TIIB[plc-tmo-mot]^WcState^WcStateIn;
                                .i_TxPDOState:=TIIB[plc-tmo-mot]^SYNC Inputs^TxPDO state;
                                '}
    plc_tmo_motion_PMPS_IO : FB_ArbiterToSubSys_IO := (RequestingSystemID := 16#F100);

    {attribute 'TcLinkTo' := '.i_RequestedBP:=TIIB[plc-tmo-optics]^IO Inputs^RequestedBP;
                                .o_CurrentBP:=TIIB[plc-tmo-optics]^IO Outputs^CurrentBP;
                                .i_Connected:=TIIB[plc-tmo-optics]^SYNC Inputs^External device not connected;
                                .i_WcState:=TIIB[plc-tmo-optics]^WcState^WcStateIn;
                                .i_TxPDOState:=TIIB[plc-tmo-optics]^SYNC Inputs^TxPDO state;
                                '}
    plc_tmo_optics_PMPS_IO : FB_ArbiterToSubSys_IO := (RequestingSystemID := 16#F101);

    {attribute 'TcLinkTo' := '.i_RequestedBP:=TIIB[plc-tmo-vac]^IO Inputs^RequestedBP;
                                .o_CurrentBP:=TIIB[plc-tmo-vac]^IO Outputs^CurrentBP;
                                .i_Connected:=TIIB[plc-tmo-vac]^SYNC Inputs^External device not connected;
                                .i_WcState:=TIIB[plc-tmo-vac]^WcState^WcStateIn;
                                .i_TxPDOState:=TIIB[plc-tmo-vac]^SYNC Inputs^TxPDO state;
                                '}
    plc_tmo_vacuum_PMPS_IO : FB_ArbiterToSubSys_IO := (RequestingSystemID := 16#F102);

    count : CTU;
//////////////////////////////////////////////
// RIX PLCs
/////////////////////////////////////////////
    {attribute 'TcLinkTo' := '.i_RequestedBP:=TIIB[plc-rix-vac]^IO Inputs^RequestedBP;
                                .o_CurrentBP:=TIIB[plc-rix-vac]^IO Outputs^CurrentBP;
                                .i_Connected:=TIIB[plc-rix-vac]^SYNC Inputs^External device not connected;
                                .i_WcState:=TIIB[plc-rix-vac]^WcState^WcStateIn;
                                .i_TxPDOState:=TIIB[plc-rix-vac]^SYNC Inputs^TxPDO state;
                                '}
    plc_rix_vac_PMPS_IO : FB_ArbiterToSubSys_IO := (RequestingSystemID := 16#F200);

    {attribute 'TcLinkTo' := '.i_RequestedBP:=TIIB[plc-rix-optics]^IO Inputs^RequestedBP;
                                .o_CurrentBP:=TIIB[plc-rix-optics]^IO Outputs^CurrentBP;
                                .i_Connected:=TIIB[plc-rix-optics]^SYNC Inputs^External device not connected;
                                .i_WcState:=TIIB[plc-rix-optics]^WcState^WcStateIn;
                                .i_TxPDOState:=TIIB[plc-rix-optics]^SYNC Inputs^TxPDO state;
                                '}
    plc_rix_optics_PMPS_IO : FB_ArbiterToSubSys_IO := (RequestingSystemID := 16#F201);

    {attribute 'TcLinkTo' := '.i_RequestedBP:=TIIB[plc-rix-mot]^IO Inputs^RequestedBP;
                                .o_CurrentBP:=TIIB[plc-rix-mot]^IO Outputs^CurrentBP;
                                .i_Connected:=TIIB[plc-rix-mot]^SYNC Inputs^External device not connected;
                                .i_WcState:=TIIB[plc-rix-mot]^WcState^WcStateIn;
                                .i_TxPDOState:=TIIB[plc-rix-mot]^SYNC Inputs^TxPDO state;
                                '}
    plc_rix_mot_PMPS_IO : FB_ArbiterToSubSys_IO := (RequestingSystemID := 16#F202);

    {attribute 'TcLinkTo' := '.i_RequestedBP:=TIIB[plc-crix-mot]^IO Inputs^RequestedBP;
                                .o_CurrentBP:=TIIB[plc-crix-mot]^IO Outputs^CurrentBP;
                                .i_Connected:=TIIB[plc-crix-mot]^SYNC Inputs^External device not connected;
                                .i_WcState:=TIIB[plc-crix-mot]^WcState^WcStateIn;
                                .i_TxPDOState:=TIIB[plc-crix-mot]^SYNC Inputs^TxPDO state;
                                '}
    plc_crix_mot_PMPS_IO : FB_ArbiterToSubSys_IO := (RequestingSystemID := 16#F203);

{attribute 'TcLinkTo' := '.i_RequestedBP:=TIIB[plc-crix-vac]^IO Inputs^RequestedBP;
                                .o_CurrentBP:=TIIB[plc-crix-vac]^IO Outputs^CurrentBP;
                                .i_Connected:=TIIB[plc-crix-vac]^SYNC Inputs^External device not connected;
                                .i_WcState:=TIIB[plc-crix-vac]^WcState^WcStateIn;
                                .i_TxPDOState:=TIIB[plc-crix-vac]^SYNC Inputs^TxPDO state;
                                '}
    plc_crix_vac_PMPS_IO : FB_ArbiterToSubSys_IO := (RequestingSystemID := 16#F205);

    {attribute 'TcLinkTo' := '.i_RequestedBP:=TIIB[plc-qrix-mot]^IO Inputs^RequestedBP;
                                .o_CurrentBP:=TIIB[plc-qrix-mot]^IO Outputs^CurrentBP;
                                .i_Connected:=TIIB[plc-qrix-mot]^SYNC Inputs^External device not connected;
                                .i_WcState:=TIIB[plc-qrix-mot]^WcState^WcStateIn;
                                .i_TxPDOState:=TIIB[plc-qrix-mot]^SYNC Inputs^TxPDO state;
                                '}


    plc_qrix_mot_PMPS_IO : FB_ArbiterToSubSys_IO := (RequestingSystemID := 16#F206);

    {attribute 'TcLinkTo' := '.i_RequestedBP:=TIIB[plc-qrix-vac]^IO Inputs^RequestedBP;
                                .o_CurrentBP:=TIIB[plc-qrix-vac]^IO Outputs^CurrentBP;
                                .i_Connected:=TIIB[plc-qrix-vac]^SYNC Inputs^External device not connected;
                                .i_WcState:=TIIB[plc-qrix-vac]^WcState^WcStateIn;
                                .i_TxPDOState:=TIIB[plc-qrix-vac]^SYNC Inputs^TxPDO state;
                                '}
    plc_qrix_vac_PMPS_IO : FB_ArbiterToSubSys_IO := (RequestingSystemID := 16#F204);

//////////////////////////////////////////////
// TXI PLCs
/////////////////////////////////////////////

    {attribute 'TcLinkTo' := '.i_RequestedBP:=TIIB[plc-txi-mot]^IO Inputs^RequestedBP;
                                .o_CurrentBP:=TIIB[plc-txi-mot]^IO Outputs^CurrentBP;
                                .i_Connected:=TIIB[plc-txi-mot]^SYNC Inputs^External device not connected;
                                .i_WcState:=TIIB[plc-txi-mot]^WcState^WcStateIn;
                                .i_TxPDOState:=TIIB[plc-txi-mot]^SYNC Inputs^TxPDO state;
                                '}
    plc_txi_motion_PMPS_IO : FB_ArbiterToSubSys_IO := (RequestingSystemID := 16#F300);

    {attribute 'TcLinkTo' := '.i_RequestedBP:=TIIB[plc-txi-optics]^IO Inputs^RequestedBP;
                                .o_CurrentBP:=TIIB[plc-txi-optics]^IO Outputs^CurrentBP;
                                .i_Connected:=TIIB[plc-txi-optics]^SYNC Inputs^External device not connected;
                                .i_WcState:=TIIB[plc-txi-optics]^WcState^WcStateIn;
                                .i_TxPDOState:=TIIB[plc-txi-optics]^SYNC Inputs^TxPDO state;
                                '}
    plc_txi_optics_PMPS_IO : FB_ArbiterToSubSys_IO := (RequestingSystemID := 16#F301);

    {attribute 'TcLinkTo' := '.i_RequestedBP:=TIIB[plc-txi-vac]^IO Inputs^RequestedBP;
                                .o_CurrentBP:=TIIB[plc-txi-vac]^IO Outputs^CurrentBP;
                                .i_Connected:=TIIB[plc-txi-vac]^SYNC Inputs^External device not connected;
                                .i_WcState:=TIIB[plc-txi-vac]^WcState^WcStateIn;
                                .i_TxPDOState:=TIIB[plc-txi-vac]^SYNC Inputs^TxPDO state;
                                '}
    plc_txi_vacuum_PMPS_IO : FB_ArbiterToSubSys_IO := (RequestingSystemID := 16#F302);

    (*Remove*)
         ar1 : bool;
 ar2 : bool;
 nReqID:UDINT;
 nReqRM:UDINT;
 bRemove:bool;
 rtRemove: R_TRIG;

END_VAR


// Updating arbiter with subsystem requests.

///////////////////////////
// KFE
    plc_kfe_motion_PMPS_IO(Arbiter:=GVL.g_fbArbiter1, fbFFHWO:=GVL.g_FastFaultOutput1, Reset:=GVL.AttemptReset, sName:= 'KFE MOTION');
    plc_kfe_vac_PMPS_IO(Arbiter:=GVL.g_fbArbiter1, fbFFHWO:=GVL.g_FastFaultOutput1, Reset:=GVL.AttemptReset, sName:= 'KFE VACUUM');
    plc_kfe_gatt_PMPS_IO(Arbiter:=GVL.g_fbArbiter1, fbFFHWO:=GVL.g_FastFaultOutput1, Reset:=GVL.AttemptReset, sName:= 'KFE GATT');
///////////////////////////

///////////////////////////
// TMO K4
// TMO-OPTICS Veto	MR1K1_IN
    plc_tmo_optics_PMPS_IO(Arbiter:=GVL.g_fbArbiter1, fbFFHWO:=GVL.g_FastFaultOutput3, Reset:=GVL.AttemptReset, sName:= 'TMO OPTICS');
// TMO-VAC and TMO-MOT OR ST3K4_IN
    plc_tmo_motion_PMPS_IO(Arbiter:=GVL.g_fbArbiter1, fbFFHWO:=GVL.g_FastFaultOutput4, Reset:=GVL.AttemptReset , sName:= 'TMO MOTION');
    plc_tmo_vacuum_PMPS_IO(Arbiter:=GVL.g_fbArbiter1, fbFFHWO:=GVL.g_FastFaultOutput4, Reset:=GVL.AttemptReset, sName:= 'TMO VACUUM');
///////////////////////////
	
//////////////////////////
// RIX
// RIX- OPTICS No Veto / Should be FFO:01 since it is upstream of all Vetos
	plc_rix_optics_PMPS_IO(Arbiter:=GVL.g_fbArbiter1, fbFFHWO:=GVL.g_FastFaultOutput1, Reset:=GVL.AttemptReset, sName:= 'RIX OPTICS');
// RIX-VAC and RIX-MOT MR1K1_OUT
    plc_rix_vac_PMPS_IO(Arbiter:=GVL.g_fbArbiter1, fbFFHWO:=GVL.g_FastFaultOutput5, Reset:=GVL.AttemptReset, sName:= 'RIX VACUUM'); 
    plc_rix_mot_PMPS_IO(Arbiter:=GVL.g_fbArbiter1, fbFFHWO:=GVL.g_FastFaultOutput5, Reset:=GVL.AttemptReset, sName:= 'RIX MOTION');
// QRIX-VAC, CRIX-VAC and CRIX-MOT MR1K1_OUT OR ST1K2_IN
	plc_crix_mot_PMPS_IO(Arbiter:=GVL.g_fbArbiter1, fbFFHWO:=GVL.g_FastFaultOutput6, Reset:=GVL.AttemptReset, sName:= 'CRIX MOTION');
    plc_crix_vac_PMPS_IO(Arbiter:=GVL.g_fbArbiter1, fbFFHWO:=GVL.g_FastFaultOutput6, Reset:=GVL.AttemptReset, sName:= 'CRIX VACUUM');
    plc_qrix_vac_PMPS_IO(Arbiter:=GVL.g_fbArbiter1, fbFFHWO:=GVL.g_FastFaultOutput6, Reset:=GVL.AttemptReset, sName:= 'QRIX VACUUM');
///////////////////////////


///////////////////////////
// TXI K3
// TXI- OPTICS No Veto / Should be FFO:01 since it is upstream of all Vetos
    plc_txi_optics_PMPS_IO(Arbiter:=GVL.g_fbArbiter1, fbFFHWO:=GVL.g_FastFaultOutput1, Reset:=GVL.AttemptReset, sName:= 'TXI OPTICS');
// TXI-VAC and TXI-MOT 	MR1K3_OUT and MR2K3_OUT
    plc_txi_vacuum_PMPS_IO(Arbiter:=GVL.g_fbArbiter1, fbFFHWO:=GVL.g_FastFaultOutput7, Reset:=GVL.AttemptReset, sName:= 'TXI VACUUM');
	plc_txi_motion_PMPS_IO(Arbiter:=GVL.g_fbArbiter1, fbFFHWO:=GVL.g_FastFaultOutput7, Reset:=GVL.AttemptReset , sName:= 'TXI MOTION');
//////////////////////////


///////////////////////////
//Beam Class override
// Dummy device for controling pmps beam parameters
fbBPControl(Arbiter:=g_fbArbiter2);

//Call the program that evaluates the Override and generate the correct Beam Parameter and adds it to arbiter 2
P_Override_Tran_BC();

////////////////////////////
// Beam parameter requestor
//////////////////////////////
fbBPRequestor(Arbiter:=GVL.g_fbArbiter2, q_ReqBP => PMPS_GVL.stRequestedBeamParameters);

//Now lets write the FAKE BP to send to the PLCs
GVL.stCurrentFakeBP := PMPS_GVL.stCurrentBeamParameters;
IF (bApplyJF) THEN
    //What if we are NOT in override mode? Then the Arbitrated1BP should be the current BP, right?
    //Should we always broadcast the requested arbitratedBP
    // yes and no. I think that it should be either the safer or the ArbitratedBP because of a specific use case in RIX OPTICS
    IF (PMPS_GVL.stCurrentBeamParameters.nTran > GVL.stArbiter1BP.nTran) THEN
        GVL.stCurrentFakeBP.nTran:= GVL.stArbiter1BP.nTran;
    END_IF
    IF (PMPS_GVL.stCurrentBeamParameters.nBeamClass > GVL.stArbiter1BP.nBeamClass) THEN
        GVL.stCurrentFakeBP.nBeamClass:= GVL.stArbiter1BP.nBeamClass;
        GVL.stCurrentFakeBP.nBCRange:= GVL.stArbiter1BP.nBCRange;
    END_IF
END_IF


// Request Cu beam rate
fbCuInterface(BP := PMPS_GVL.stRequestedBeamParameters);


// Keep an eye on the photon energy
fbPhotonEnergyWatcher(i_stCurrentBeamParams	:= PMPS_GVL.stCurrentBeamParameters,
                    i_stRequestedBeamParams := PMPS_GVL.stRequestedBeamParameters,
                    io_fbFFHWO:= GVL.g_FastFaultOutput1,
                    i_xReset := GVL.AttemptReset);

//Assert beam class
P_BeamClassAssertion();


//Use Only in very critical cases. Only when you are sure. This might result in damage to devices
(*remove*)
(*Debugging functions*)
ar1:= GVL.g_fbArbiter1.CheckRequestInPool(nReqRM);

rtRemove(CLK:= bRemove);
if (rtRemove.Q) THEN
     GVL.g_fbArbiter1.RemoveRequest(nReqRM);
END_IF

END_PROGRAM

// ---- POUs/TEMP/FB_ArbiterToSubSys_IO.TcPOU
(* Exchanges preemption requests and current beam state with subsystems in arbiter
network.

2019-12-2, A. Wallace

Use in conjunction with FB_SubSysToArbiter_IO.

This FB runs in the beamline arbiter PLC (BAP). There should be one of these for every
subsystem interfaced to the BAP. Each subsystem PLC should run a sibling FB_SubSysToArbiter_IO FB.

This FB and its subordinate communicate through the ethercat connection between the subsystem PLC and the BAP.

A beam parameter set request is sent from the subsystem to this PLC, and includes a cohort number.

This cohort number (i_RequestedBP.nCohortInt) is compared to a local cohort number (nRequestedCohort).
A request from the subsystem to update or modify its current request is indicated by an increase in the
i_RequestedBP.nCohortInt value. Then this function block updates the local arbiter request for the subsystem
and awaits confirmation. Once the new request is confirmed in the preemptive system this function block increments
the ActiveCohort value to match the nRequestedCohort. ActiveCohort is also relayed back to the subsystem
as the active cohort value in the o_CurrentBP set. The subsystem then knows its request has been heard,
and can carry out its own acknowledgement to its various requestors.

Things to note:
If a subsystem has any new or changed preemptive requests you should see the cohort value increment a bit.
If the cohort number is incrementing out of control, it usually means the subsysetm has some preemptive
request loop (two arbiters elevating to each other), or there is a RequestAdd, RequestRemove loop.

*)
FUNCTION_BLOCK FB_ArbiterToSubSys_IO
VAR_INPUT
    RequestingSystemID	:	DWORD := PMPS_GVL.EXCLUDED_ASSERTION_ID; // System ID for making requests to the supreme arbiter
    sName : STRING := 'ArbiterToSubSys';
    Reset : BOOL;
END_VAR
VAR_OUTPUT
END_VAR
VAR_IN_OUT
    Arbiter	: FB_Arbiter;
    fbFFHWO : FB_HardwareFFOutput;
END_VAR
VAR

    i_RequestedBP AT %I*	:	ST_BeamParams_IO; // Requested BP from subsystem
    {attribute 'pytmc' := '
        pv: RequestedBP:FromSubSys
    '}
    RequestedBP: ST_BeamParams;

    o_CurrentBP AT %Q* : ST_BeamParams_IO; // Current BP set

    // EL6692 Diagnostics
    i_Connected AT %I* : BOOL; // SYNC Inputs^External device not connected !!! Doesn't really work.
    {attribute 'pytmc' := 'pv: WcState
        io: i
        field: DESC Working counter state.
        field: ZNAM OK
        field: ONAM Error'}
    i_WcState AT %I* : BOOL := TRUE; // WcState^WcState
    {attribute 'pytmc' := 'pv: TxPDO_state
        io: i
        field: DESC PDO Transmission is OK
        field: ZNAM OK
        field: ONAM Error'}
    i_TxPDOState AT %I* : BOOL := TRUE; // SYNC Inputs^TxPDO state
    {attribute 'pytmc' := 'pv: TxPDO_toggle
        io: i
        field: DESC PDO Transmission is OK
        field: ZNAM OK
        field: ONAM Error'}
    i_TxPDOToggle AT %I* : BOOL; // TxPDO toggle

    // Fast faults
    ffPMPSIO_Disconnect : FB_FastFault := (i_Desc:='Issue w/ arbiter interface to subsystem, verify subsystem is OK, or ethercat connection.'); // Fast fault for ethercat issues
    nActiveCohort : UDINT := 0; // Active cohort. Updated to the req. number from the sub system after request is confirmed.
    nRequestedCohort : UDINT := 0;
    rtToggle : R_TRIG;


END_VAR


// Incoming request from subsystem PLC
RequestedBP := IO_TO_BP(i_RequestedBP);

// Update Arbiter with our request
rtToggle(CLK:= i_RequestedBP.xValid); // If interface resumes, reset/catch up
// xValid will go false if the PLC program on the other side is stopped. Ironically the ethercat interface continues happily.
// If subsystem cohort has incremented, update beam parameter request with our arbiter
IF rtToggle.Q THEN
    nActiveCohort := 0;
END_IF

IF i_RequestedBP.nCohortInt > nRequestedCohort OR rtToggle.Q THEN
    Arbiter.RemoveRequest(RequestingSystemID);
    Arbiter.AddRequest(RequestingSystemID, RequestedBP,sName);
    nRequestedCohort := i_RequestedBP.nCohortInt;
END_IF


// Check if latest request is acknowledged by this arbiter
// Acknowledgement happens after an arbitration cycle, which means if RequestedCohort just incremented
// due to a new request, CheckRequest will be false.
IF Arbiter.CheckRequest(RequestingSystemID) THEN
    nActiveCohort := nRequestedCohort; // If it is, then the active cohort is set to the requested cohort number.
END_IF

// Sending current beam parameter set to subsystems
o_CurrentBP := BP_TO_IO(GVL.stCurrentFakeBP);//MG: Not Sure, the Idea it is the Current but with fake transmission and Beamclass??
o_CurrentBP.nCohortInt := nActiveCohort;


//////////////////////////////////////
// Verifying the ethercat interface health
/////////////////////////////////////
// Both of these values should be 0 for a fully valid exchange
ffPMPSIO_Disconnect.i_xOK := NOT i_WcState AND NOT i_TxPDOState;

ffPMPSIO_Disconnect(
    io_fbFFHWO := fbFFHWO,
    i_xReset := Reset,
    i_DevName := sName,
    i_TypeCode:=5);

END_FUNCTION_BLOCK

// ---- POUs/P_Override_Tran_BC.TcPOU
PROGRAM P_Override_Tran_BC
VAR
    fbBPRequestor_Arbiter1 : FB_BPRequestor; // gets the arbiter 1 BP
    stOverrideBP:ST_BeamParams;
    stPreviousOverrideBP:ST_BeamParams;
    tDuration:TIME;
    tonDuration:TON;
    {attribute 'pytmc' := '
       pv: @(PREFIX)RequestedPowerMax
    '}
    rPowerMax:REAL;
    {attribute 'pytmc' := '
       pv: @(PREFIX)PowerOverride
    '}
    rPowerOverride:REAL;
    arrTableBC	: ARRAY[1..16,1..2] OF REAL;
    arrIndex: INT;
    bInit : BOOl:= TRUE;
END_VAR

IF bInit THEN
    ACT_INIT(); // not needed every cycle
    bInit := FALSE;
END_IF


//Beam intensity factor implemenation
// No diff by zero
IF (nBeamIntensityJF =0) OR (nBeamIntensityJF > GVL.nBeamIntensity ) THEN nBeamIntensityJF:=GVL.nBeamIntensity; END_IF
//Check it it has expired or is cancelled and reset to defaults
IF(tonDuration.Q OR bCancelJF)
THEN
    nBeamIntensityJF:=GVL.nBeamIntensity;
    bCancelJF := FALSE;
     bApplyJF := FALSE;
END_IF

//Get the Beam paramters from Arbiter 1
fbBPRequestor_Arbiter1(Arbiter:=GVL.g_fbArbiter1, q_ReqBP =>stArbiter1BP);
//Start with Override to be equal to the Arbiter1 Beam parameters
stOverrideBP := stArbiter1BP;

// Maximum duration is 12 hours
rDurationJF := LIMIT(0,rDurationJF,MaxDuration);
//check if it is applied
tDuration:= TO_TIME(rDurationJF*60*60*1000);//to msec
tonDuration(IN:=bApplyJF,PT:=tDuration,ET=>);
rTimeRemainJF:= rDurationJF - (TO_REAL(tonDuration.ET)/60/60/1000);//to hours


 // Send request from this arbiter to the gas attenuator
 IF (bApplyJF) THEN
     //Transmission override
      stOverrideBP.nTran := LIMIT(0,(GVL.nBeamIntensity/nBeamIntensityJF)*stArbiter1BP.nTran*PMPS_GVL.TRANS_SCALING_FACTOR,1);
     // Beamclass override
     arrIndex := stArbiter1BP.nBeamClass+1;
     //Make sure to remain within the bounds of the array
     arrIndex := LIMIT(1,arrIndex,16);
     //Look up the Max power for this beamclass
     rPowerMax := arrTableBC[arrIndex,2];
     //Calculate the new max allowed power based on the current beam class power and judgement factor
     rPowerOverride:= ((GVL.nBeamIntensity/nBeamIntensityJF)*stArbiter1BP.nTran)*rPowerMax;
     //If Power override is lower Than Power Max, keep Power Max
     IF ( rPowerOverride < rPowerMax) THEN rPowerOverride := rPowerMax; END_IF
     //Look up the new beamclass for the adjusted power
     stOverrideBP.nBeamClass := TO_USINT(M_LookUp(rPowerOverride,arrTableBC));
     // Apply bitmask to BC range
     stOverrideBP.nBCRange:= SHL(1,stOverrideBP.nBeamClass)-1;
END_IF

// Add the override BP to arbiter 2, so it is arbitrated with the beamline parameter
IF F_DifferentBeamParams (stPreviousOverrideBP,stOverrideBP) THEN
    GVL.g_fbArbiter2.RemoveRequest(16#FFF1);
    GVL.g_fbArbiter2.AddRequest(nReqID := 16#FFF1, stReqBp := stOverrideBP, sDevName := 'Beamlines Summary');
    stPreviousOverrideBP := stOverrideBP;
END_IF

ACTION ACT_Init:
IF bInit
THEN
    (* init array with BeamClass Data  *)
    (* 	BeamClass		 |		Power		*)
    arrTableBC[1,1] := 0;	arrTableBC[1,2] := 0;
    arrTableBC[2,1] := 1;	arrTableBC[2,2] := 0;
    arrTableBC[3,1] := 2;	arrTableBC[3,2] := 1.4;
    arrTableBC[4,1] := 3;	arrTableBC[4,2] := 14;
    arrTableBC[5,1] := 4;	arrTableBC[5,2] := 40;
    arrTableBC[6,1] := 5;	arrTableBC[6,2] := 60;
    arrTableBC[7,1] := 6;	arrTableBC[7,2] := 140;
    arrTableBC[8,1] := 7;	arrTableBC[8,2] := 1200;
    arrTableBC[9,1] := 8;	arrTableBC[9,2] := 6000;
    arrTableBC[10,1] := 9;	arrTableBC[10,2] := 12000;
    arrTableBC[11,1] := 10;	arrTableBC[11,2] := 30000;
    arrTableBC[12,1] := 11; arrTableBC[12,2] := 60000;
    arrTableBC[13,1] := 12;	arrTableBC[13,2] := 120000;
    arrTableBC[14,1] := 13;	arrTableBC[14,2] := 120000;
    arrTableBC[15,1] := 14;	arrTableBC[15,2] := 120000;
    arrTableBC[16,1] := 15;	arrTableBC[16,2] := 120000;

    bInit:=False;

END_IF
END_ACTION

METHOD M_LookUp : REAL
VAR_INPUT
    Pnew : LREAL;
    arrTableBC	: ARRAY[1..16,1..2] OF REAL;
END_VAR

VAR
    iIndex: INT;
END_VAR

VAR CONSTANT
    iLowBound :INT :=1;
    iHighBound:INT :=16;
END_VAR
M_LookUp:=0;
FOR iIndex := iLowBound TO iHighBound DO
    (*Need to avoid Floating-Point Comparison issue*)
    // Ceiling function isn't available for this build only available on TwinCAT v3.1 >= 4026.13
    IF (FLOOR(Pnew)+ 1 >= arrTableBC[iIndex,2]) THEN M_LookUp := arrTableBC[iIndex,1];
        ELSE return;
    END_IF
END_FOR
END_METHOD

END_PROGRAM

// ---- POUs/P_BeamClassAssertion.TcPOU
PROGRAM P_BeamClassAssertion
VAR
    {attribute 'pytmc' := '
    pv: @(PREFIX)BeamClassWatcher
    '}
    fbBeamClassWatcher : FB_BeamClassWatcher;
    {attribute 'pytmc' := '
    pv: @(PREFIX)BeamClassOutputs
    '}
    fbMPSInterface	:	FB_BeamClassOutputs_BCD;

END_VAR


// Request beam class
fbMPSInterface(BP := PMPS_GVL.stRequestedBeamParameters);

// Keep an eye on the beam class
fbBeamClassWatcher(i_stCurrentBeamParams	:= PMPS_GVL.stCurrentBeamParameters,
                    i_stRequestedBeamParams := PMPS_GVL.stRequestedBeamParameters,
                    io_fbFFHWO:= GVL.g_FastFaultOutput1,
                    i_xAutoReset := TRUE);

END_PROGRAM

// ---- POUs/P_AT1K0_SL1K0.TcPOU
PROGRAM P_AT1K0_SL1K0
VAR

    // Transmisison request and status with plc-kfe-gatt
    {attribute 'TcLinkTo' := 'TIIB[plc-kfe-gatt]^IO Outputs^Requested Transmission'}
    q_nTranToAT1K0Req AT %Q* : ST_PMPS_Attenuator_IO; // Transmission request to AT1K0
    {attribute 'TcLinkTo' := 'TIIB[plc-kfe-gatt]^IO Inputs^Current Transmission'}
    i_nTranToAT1K0Stat AT %I* : ST_PMPS_Attenuator_IO; // Transmission request to AT1K0

    // plc-kfe-gatt interface diagnostics
    {attribute 'TcLinkTo' := 'TIIB[plc-kfe-gatt]^WcState^WcStateOut'}
    i_bWcStateOut_AT1K0 AT %I* : BOOL;
    {attribute 'TcLinkTo' := 'TIIB[plc-kfe-gatt]^WcState^WcStateIn'}
    i_bWcStateIn_AT1K0 AT %I* : BOOL;
    {attribute 'TcLinkTo' := 'TIIB[plc-kfe-gatt]^InfoData^State'}
    i_nState_AT1K0 AT %I* : UINT;

    // Apterure request and status to plc-kfe-motion
    {attribute 'TcLinkTo' := 'TIIB[plc-kfe-motion]^IO Outputs^AptArrayReq'}
    q_stAptArrayReq AT %Q* : ARRAY [1..4] OF ST_PMPS_Aperture_IO;
    {attribute 'TcLinkTo' := 'TIIB[plc-kfe-motion]^IO Inputs^AptArrayStatus'}
    i_stAptArrayStat AT %I* : ARRAY [1..4] OF ST_PMPS_Aperture_IO;

    // plc-kfe-motion interface diagnostics
    {attribute 'TcLinkTo' := 'TIIB[plc-kfe-motion]^WcState^WcStateOut'}
    i_bWcStateOut_KFEMOT AT %I* : BOOL;
    {attribute 'TcLinkTo' := 'TIIB[plc-kfe-motion]^WcState^WcStateIn'}
    i_bWcStateIn_KFEMOT AT %I* : BOOL;
    {attribute 'TcLinkTo' := 'TIIB[plc-kfe-motion]^InfoData^State'}
    i_nState_KFEMOT AT %I* : UINT;

    idx : UINT;

    ffKFEMotConnection : FB_FastFault := (
        i_DevName := 'PMPS Arbiter',
        i_Desc := 'EtherCAT interface watcher, for connection to KFE Motion systems for SL1K0 size requests. Very rare. Make a note, and if it can be reset, go ahead.',
        i_TypeCode := 16#5);
    ffKFEGattConnection : FB_FastFault := (
        i_DevName := 'PMPS Arbiter',
        i_Desc := 'EtherCAT interface watcher, for connection to KFE Gas Att. systems for Transmission requests. Very rare. Make a note, and if it can be reset, go ahead.',
        i_TypeCode := 16#5);
    bSimApt: BOOL;

    tDuration:TIME;
    tonDuration:TON;


END_VAR


// If interface with plc-kfe-gatt OK carry out exchange
IF i_bWcStateOut_AT1K0 = 0 AND i_bWcStateIn_AT1K0 = 0 AND i_nState_AT1K0 = 8 THEN
    q_nTranToAT1K0Req.nTran := PMPS_GVL.stRequestedBeamParameters.nTran*PMPS_GVL.TRANS_SCALING_FACTOR;
    PMPS_GVL.stCurrentBeamParameters.nTran := i_nTranToAT1K0Stat.nTran;
    q_nTranToAT1K0Req.xAttOK := 16#FF;
    ffKFEGattConnection.i_xOK := TRUE;
ELSE
    // Fast fault
    ffKFEGattConnection.i_xOK := FALSE;
    PMPS_GVL.stCurrentBeamParameters.nTran := PMPS_GVL.TRANS_SCALING_FACTOR;//100;

END_IF

ffKFEGattConnection(io_fbFFHWO := g_FastFaultOutput1);

// If interface with plc-kfe-motion OK, carry out exchange
IF i_bWcStateIn_KFEMOT = 0 AND i_bWcStateOut_KFEMOT = 0 AND i_nState_KFEMOT = 8 THEN

    // Send request from this arbiter to kfe-mot
    MEMCPY( ADR(q_stAptArrayReq) , ADR(PMPS_GVL.stRequestedBeamParameters.astApertures) , PMPS_GVL.MAX_APERTURES * SIZEOF(ST_PMPS_Aperture_IO) );

    // 	Recieve current apreture state for broadcast
    MEMCPY( ADR(PMPS_GVL.stCurrentBeamParameters.astApertures) , ADR(i_stAptArrayStat) , PMPS_GVL.MAX_APERTURES * SIZEOF(ST_PMPS_Aperture_IO) );

    ffKFEMotConnection.i_xOK := TRUE;

ELSIF bSimApt THEN
    PMPS_GVL.stCurrentBeamParameters.astApertures := PMPS_GVL.stRequestedBeamParameters.astApertures;
ELSE
    // Fast fault
    ffKFEMotConnection.i_xOK := FALSE;
    // Set broadcast apterture states to not OK
    FOR idx := 1 TO PMPS_GVL.MAX_APERTURES DO
        PMPS_GVL.stCurrentBeamParameters.astApertures[idx].xOK := FALSE;
    END_FOR
END_IF

ffKFEMotConnection(io_fbFFHWO := g_FastFaultOutput1);

END_PROGRAM

// ---- POUs/P_SATT.TcPOU
PROGRAM P_SATT
VAR
    //All Sold attenuators requests are summerrized into this one output
    q_SattArrayReq AT %Q* : ARRAY [1..PMPS_GVL.AUX_ATTENUATORS] OF ST_PMPS_Attenuator_IO; // Transmission request to ALL PLCs
    //Per PLC current satt trans
    {attribute 'TcLinkTo' := 'TIIB[plc-kfe-motion]^IO Inputs^SattArrayStatus'}
    i_SattArrayStatus_KFE AT %I* : ARRAY [1..PMPS_GVL.AUX_ATTENUATORS] OF ST_PMPS_Attenuator_IO; // Transmission request to KFE MOT PLC
        {attribute 'TcLinkTo' := 'TIIB[plc-rix-mot]^IO Inputs^SattArrayStatus'}
    i_SattArrayStatus_RIX AT %I* : ARRAY [1..PMPS_GVL.AUX_ATTENUATORS] OF ST_PMPS_Attenuator_IO; // Transmission request to RIX MOT PLC

    // plc-tmo-mot interface diagnostics
    {attribute 'TcLinkTo' := 'TIIB[plc-kfe-motion]^WcState^WcStateOut'}
    i_bWcStateOut_kfe_mot AT %I* : BOOL;
    {attribute 'TcLinkTo' := 'TIIB[plc-kfe-motion]^WcState^WcStateIn'}
    i_bWcStateIn_kfe_mot AT %I* : BOOL;
    {attribute 'TcLinkTo' := 'TIIB[plc-kfe-motion]^InfoData^State'}
    i_nState_kfe_mot AT %I* : UINT;

    // plc-rix-mot interface diagnostics
    {attribute 'TcLinkTo' := 'TIIB[plc-rix-mot]^WcState^WcStateOut'}
    i_bWcStateOut_rix_mot AT %I* : BOOL;
    {attribute 'TcLinkTo' := 'TIIB[plc-rix-mot]^WcState^WcStateIn'}
    i_bWcStateIn_rix_mot AT %I* : BOOL;
    {attribute 'TcLinkTo' := 'TIIB[plc-rix-mot]^InfoData^State'}
    i_nState_rix_mot AT %I* : UINT;

    //FFO Connection per PLC
    ffkfeConnection : FB_FastFault := (
        i_DevName := 'PMPS Arbiter',
        i_Desc := 'EtherCAT interface watcher, for tmo-mot connection to systems for attenuation requests. Very rare. Make a note, and if it can be reset, go ahead.',
        i_TypeCode := 16#5);
    ffRixConnection : FB_FastFault := (
        i_DevName := 'PMPS Arbiter',
        i_Desc := 'EtherCAT interface watcher, for rix-mot connection to systems for attenuation requests. Very rare. Make a note, and if it can be reset, go ahead.',
        i_TypeCode := 16#5);
END_VAR



// Send request from this arbiter to all satts
MEMCPY( ADR(q_SattArrayReq) , ADR(PMPS_GVL.stRequestedBeamParameters.astAttenuators) , PMPS_GVL.AUX_ATTENUATORS * SIZEOF(ST_PMPS_Attenuator_IO) );

//TMO motion PLC SATT current trans update
IF i_bWcStateIn_kfe_mot = 0 AND i_bWcStateOut_kfe_mot = 0 AND i_nState_kfe_mot = 8 THEN
    // 	Recieve current transmission of the satt
    //PMPS_GVL.stCurrentBeamParameters.astAttenuators[PMPS.K_Attenuators.AT1K4].nTran :=  i_SattArrayStatus_KFE[PMPS.K_Attenuators.AT1K4].nTran;
    //PMPS_GVL.stCurrentBeamParameters.astAttenuators[PMPS.K_Attenuators.AT1K4].xAttOK :=  i_SattArrayStatus_KFE[PMPS.K_Attenuators.AT1K4].xAttOK;
    ffkfeConnection.i_xOK := TRUE;
ELSE
    // Fast fault
    ffkfeConnection.i_xOK := FALSE;
END_IF
ffkfeConnection(io_fbFFHWO := g_FastFaultOutput1);

//RIX motion PLC SATT current trans update
IF i_bWcStateIn_rix_mot = 0 AND i_bWcStateOut_rix_mot = 0 AND i_nState_rix_mot = 8 THEN

    // 	Recieve current transmission of the satt
    //PMPS_GVL.stCurrentBeamParameters.astAttenuators[PMPS.K_Attenuators.AT1K2].nTran :=  i_SattArrayStatus_RIX[PMPS.K_Attenuators.AT1K2].nTran;
    //PMPS_GVL.stCurrentBeamParameters.astAttenuators[PMPS.K_Attenuators.AT1K2].xAttOK :=  i_SattArrayStatus_RIX[PMPS.K_Attenuators.AT1K2].xAttOK;
    //PMPS_GVL.stCurrentBeamParameters.astAttenuators[PMPS.K_Attenuators.AT2K2].nTran :=  i_SattArrayStatus_RIX[PMPS.K_Attenuators.AT2K2].nTran;
    //PMPS_GVL.stCurrentBeamParameters.astAttenuators[PMPS.K_Attenuators.AT2K2].xAttOK :=  i_SattArrayStatus_RIX[PMPS.K_Attenuators.AT2K2].xAttOK;
    ffRixConnection.i_xOK := TRUE;
ELSE
    // Fast fault
    ffRixConnection.i_xOK := FALSE;
END_IF
ffRixConnection(io_fbFFHWO := g_FastFaultOutput1);

END_PROGRAM

// ---- POUs/Fast_Faults_Evaluate.TcPOU
PROGRAM Fast_Faults_Evaluate
VAR
FFO    :    FB_FastFault :=(i_DevName := 'PMPS Arbiter',
        i_Desc := 'Fault occurs when the beamline valves on qrixs are not in open state',
        i_TypeCode := 16#1010);
i_xFastFaultOut_qrix_vac AT %I*:        BOOL;

FFO2   :    FB_FastFault :=(i_DevName := 'PMPS Arbiter',
        i_Desc := 'Forward Fault from TXI Vacuum.',
        i_TypeCode := 16#3010);
 {attribute 'TcLinkTo' := 'TIIB[plc-txi-vac]^IO Inputs^FFO'}
i_xFastFaultOut_txi_vac AT %I*:        BOOL;

FFO3    :    FB_FastFault :=(i_DevName := 'PMPS Arbiter',
        i_Desc := 'Forward Fault from TXI Motion.',
        i_TypeCode := 16#3013);
{attribute 'TcLinkTo' := 'TIIB[plc-txi-mot]^IO Inputs^FFO'}
i_xFastFaultOut_txi_mot AT %I*:        BOOL;


FFO4    :    FB_FastFault :=(i_DevName := 'PMPS Arbiter',
        i_Desc := 'Forward Fault from TXI OPTICS.',
        i_TypeCode := 16#3013);
{attribute 'TcLinkTo' := 'TIIB[plc-txi-optics]^IO Inputs^FFO'}
i_xFastFaultOut_txi_optics AT %I*:        BOOL;

(*TXI OPTICS Protection Faults*)

FFO_RIX_TXI_OPTICS :    FB_FastFault :=(i_DevName := 'PMPS Arbiter',
        i_Desc := 'Fault when MR1K1 and/or K3 mirrors are in inconsistent state',
        i_TypeCode := 16#3103);

FFO_TXI_OPTICS :    FB_FastFault :=(i_DevName := 'PMPS Arbiter',
        i_Desc := 'Fault when MR1K3 is OUT and MR2K3 is IN',
        i_TypeCode := 16#3113);
// This is to link 3,4,5,6,7 to an actual cactive fault 2
FFO34567to2link :    FB_FastFault :=(i_DevName := 'Hutch PLC Communication',
        i_Desc := 'Hutch PLC to Arbiter communication error, please check faults below',
        i_TypeCode := 16#00C0);

// This is an RP required FFO
RP_HighBeamPower :    FB_FastFault :=(i_DevName := 'HighPowerBeam fault',
        i_Desc := 'High power beam not allowed to terminate in the FEE',
        i_TypeCode := 16#5AFE);
END_VAR

//RQRIX Forard Fault
FFO(
    io_fbFFHWO := g_FastFaultOutput6,
    i_xOK := i_xFastFaultOut_qrix_vac,
    i_xAutoReset := TRUE);

//TXI Forward Faults
FFO2(
    io_fbFFHWO := g_FastFaultOutput7,
    i_xOK := i_xFastFaultOut_txi_vac,
    i_xAutoReset := TRUE);

FFO3(
    io_fbFFHWO := g_FastFaultOutput7,
    i_xOK := i_xFastFaultOut_txi_mot,
    i_xAutoReset := TRUE);

FFO4(
    io_fbFFHWO := g_FastFaultOutput1,
    i_xOK := i_xFastFaultOut_txi_optics,
    i_xAutoReset := TRUE);


(*TXI OPTICS Protection Faults*)
(* MR1K1 | MR1K3 | MR2K3 | Fault *)
(*  IN   |  IN   |  OUT  | TRUE  *)
(*  IN   |  OUT  |  IN   | TRUE  *)
(*  IN   |  IN   |  IN   | TRUE  *)
(*  OUT  |  IN   |  OUT  | TRUE  *)
(*  OUT  |  OUT  |  IN   | TRUE  *)

FFO_RIX_TXI_OPTICS(
    io_fbFFHWO := g_FastFaultOutput1,
    i_xOK := (PMPS_GVL.stCurrentBeamParameters.aVetoDevices[PMPS.K_Stopper.MR1K1_IN] AND NOT PMPS_GVL.stCurrentBeamParameters.aVetoDevices[PMPS.K_Stopper.MR1K1_OUT])
                AND ((PMPS_GVL.stCurrentBeamParameters.aVetoDevices[PMPS.K_Stopper.MR1K3_OUT] AND NOT PMPS_GVL.stCurrentBeamParameters.aVetoDevices[PMPS.K_Stopper.MR1K3_IN])
                    AND (PMPS_GVL.stCurrentBeamParameters.aVetoDevices[PMPS.K_Stopper.MR2K3_OUT] AND NOT PMPS_GVL.stCurrentBeamParameters.aVetoDevices[PMPS.K_Stopper.MR2K3_IN]))
                OR (PMPS_GVL.stCurrentBeamParameters.aVetoDevices[PMPS.K_Stopper.MR1K1_OUT] AND NOT PMPS_GVL.stCurrentBeamParameters.aVetoDevices[PMPS.K_Stopper.MR1K1_IN]) ,
    i_xAutoReset := TRUE);

FFO_TXI_OPTICS(
    io_fbFFHWO := g_FastFaultOutput1,
    i_xOK := (PMPS_GVL.stCurrentBeamParameters.aVetoDevices[PMPS.K_Stopper.MR1K3_OUT] AND NOT PMPS_GVL.stCurrentBeamParameters.aVetoDevices[PMPS.K_Stopper.MR1K3_IN]
                    AND PMPS_GVL.stCurrentBeamParameters.aVetoDevices[PMPS.K_Stopper.MR2K3_OUT] AND NOT PMPS_GVL.stCurrentBeamParameters.aVetoDevices[PMPS.K_Stopper.MR2K3_IN])
                OR (PMPS_GVL.stCurrentBeamParameters.aVetoDevices[PMPS.K_Stopper.MR1K3_IN] AND NOT PMPS_GVL.stCurrentBeamParameters.aVetoDevices[PMPS.K_Stopper.MR1K3_OUT]
                    AND PMPS_GVL.stCurrentBeamParameters.aVetoDevices[PMPS.K_Stopper.MR2K3_IN] AND NOT PMPS_GVL.stCurrentBeamParameters.aVetoDevices[PMPS.K_Stopper.MR2K3_OUT])  ,
    i_xAutoReset := TRUE);

FFO34567to2link(
	  io_fbFFHWO := g_FastFaultOutput2,
	   i_xOK := g_FastFaultOutput3.q_xFastFaultOut AND g_FastFaultOutput4.q_xFastFaultOut AND g_FastFaultOutput5.q_xFastFaultOut AND g_FastFaultOutput6.q_xFastFaultOut AND g_FastFaultOutput7.q_xFastFaultOut ,
       i_xAutoReset := TRUE);
	
// RP requested fault
RP_HighBeamPower(
io_fbFFHWO := g_FastFaultOutput1,
i_xOK := ((PMPS_GVL.stCurrentBeamParameters.nBeamClass >9 AND PMPS_GVL.stCurrentBeamParameters.nTran >=0.4) (*High Power Beam*)
             AND ((PMPS_GVL.stCurrentBeamParameters.aVetoDevices[PMPS.K_Stopper.MR1K1_OUT] AND NOT PMPS_GVL.stCurrentBeamParameters.aVetoDevices[PMPS.K_Stopper.ST3K4]) (* Beam in TMO*)
               OR (PMPS_GVL.stCurrentBeamParameters.aVetoDevices[PMPS.K_Stopper.MR1K1_IN] AND  NOT PMPS_GVL.stCurrentBeamParameters.aVetoDevices[PMPS.K_Stopper.ST1K2]))) (*BEAM in RIX*)
            OR (PMPS_GVL.stCurrentBeamParameters.nBeamClass<=9)(*LOW Power Beam *)
            OR ((PMPS_GVL.stCurrentBeamParameters.nBeamClass>=9) AND (PMPS_GVL.stCurrentBeamParameters.nTran <0.4))
            OR PMPS_GVL.stCurrentBeamParameters.nMachineMode = 0, // Machine is running in NC mode
i_xAutoReset := FALSE);

//Execute /evaulate FFOs
// Evaluate fast fault No Vetos
g_FastFaultOutput1.Execute();
g_FastFaultOutput2.EvaluateOutput(bAutoReset:=TRUE);
// Evaluate fast fault vetos TMO
//TMO-OPTICS Veto	MR1K1_IN
g_FastFaultOutput3.Execute(i_xVeto:= PMPS_GVL.stCurrentBeamParameters.aVetoDevices[PMPS.K_Stopper.MR1K1_IN],bAutoReset:=TRUE);
// TMO-VAC and TMO-MOT ST3K4_IN
g_FastFaultOutput4.Execute(i_xVeto:= PMPS_GVL.stCurrentBeamParameters.aVetoDevices[PMPS.K_Stopper.ST3K4],bAutoReset:=TRUE);
// Evaluate fast fault vetos RIX
// RIX-VAC and RIX-MOT MR1K1_OUT
g_FastFaultOutput5.Execute(i_xVeto:= PMPS_GVL.stCurrentBeamParameters.aVetoDevices[PMPS.K_Stopper.MR1K1_OUT],bAutoReset:=TRUE);
// QRIX-VAC, CRIX-VAC and CRIX-MOT MR1K1_OUT OR ST1K2_IN
g_FastFaultOutput6.Execute(i_xVeto:= PMPS_GVL.stCurrentBeamParameters.aVetoDevices[PMPS.K_Stopper.MR1K1_OUT] OR PMPS_GVL.stCurrentBeamParameters.aVetoDevices[PMPS.K_Stopper.ST1K2],bAutoReset:=TRUE);
// Evaluate fast fault vetos TXI
// TXI-VAC and TXI-MOT 	MR1K3_OUT and MR2K3_OUT
g_FastFaultOutput7.Execute(i_xVeto:= PMPS_GVL.stCurrentBeamParameters.aVetoDevices[PMPS.K_Stopper.MR1K3_OUT] AND PMPS_GVL.stCurrentBeamParameters.aVetoDevices[PMPS.K_Stopper.MR2K3_OUT],bAutoReset:=TRUE);

END_PROGRAM

// ---- POUs/Testing.TcPOU
PROGRAM Testing
VAR
    AttemptReset : TON := (PT:=T#1s);
    gAttemptReset : TON := (PT:=T#500ms);

    testFF : FB_FastFault;
    cycle : INT;
END_VAR


// Trip a fast fault periodically
testFF(io_fbFFHWO:= g_FastFaultOutput1);
//testFF.i_xOK := (cycle mod 1000) = 0;
//cycle := cycle + 1;

//Periodically try to reset the photon energy fault.
AttemptReset(IN:=PMPS_Arbiter.fbPhotonEnergyWatcher.xPhotonEnergyWithinBounds, Q=>GVL.AttemptReset);

gAttemptReset(IN:=GVL.g_FastFaultOutput1.xOK, Q=>GVL.g_FastFaultOutput1.i_xReset);

END_PROGRAM

// ---- ImplicitChecks/CheckBounds.TcPOU
// Implicitly generated code : DO NOT EDIT
FUNCTION CheckBounds : DINT
VAR_INPUT
    index, lower, upper: DINT;
END_VAR
// User defined local variables
VAR
    sMessageLow   : STRING := 'CheckBounds: Index too low (%d)';
    sMessageHigh  : STRING := 'CheckBounds: Index too high (%d)';
END_VAR

// Index too low
IF index < lower THEN
    CheckBounds := lower;
    // Increase global counter
    GVL_CheckBounds.nTooLow := GVL_CheckBounds.nTooLow + 1;
    // Log message
    ADSLOGDINT(msgCtrlMask := ADSLOG_MSGTYPE_WARN,
               msgFmtStr   := sMessageLow,
               dintArg     := index);

// Index too high
ELSIF index > upper THEN
    CheckBounds := upper;
    // Increase global counter
    GVL_CheckBounds.nTooHigh := GVL_CheckBounds.nTooHigh + 1;
    // Log message
    ADSLOGDINT(msgCtrlMask := ADSLOG_MSGTYPE_WARN,
               msgFmtStr   := sMessageHigh,
               dintArg     := index);

// Index OK
ELSE
    CheckBounds := index;
END_IF
{flow}

END_FUNCTION

// ---- ImplicitChecks/CheckRangeSigned.TcPOU
// Implicitly generated code : DO NOT EDIT
FUNCTION CheckRangeSigned : DINT
VAR_INPUT
    value, lower, upper: DINT;
END_VAR

// Implicitly generated code : Only an Implementation suggestion

IF (value < lower) THEN
    CheckRangeSigned := lower;
ELSIF(value > upper) THEN
    CheckRangeSigned := upper;
ELSE
    CheckRangeSigned := value;
END_IF
{flow}

END_FUNCTION

// ---- ImplicitChecks/CheckRangeUnsigned.TcPOU
// Implicitly generated code : DO NOT EDIT
FUNCTION CheckRangeUnsigned : UDINT
VAR_INPUT
    value, lower, upper: UDINT;
END_VAR

// Implicitly generated code : Only an Implementation suggestion
{noflow}
IF (value < lower) THEN
    CheckRangeUnsigned := lower;
ELSIF(value > upper) THEN
    CheckRangeUnsigned := upper;
ELSE
    CheckRangeUnsigned := value;
END_IF
{flow}

END_FUNCTION

// ---- POUs/CXDisplay.TcPOU
PROGRAM CXDisplay
VAR
    DisplayStats : FB_CXSetTextDisplayUSB := (nPort:=28928);
    fbFormat   : FB_FormatString;
    bError     : BOOL;
    nErrID     : UDINT;
    sOut       : T_MaxString;
END_VAR

(*
DisplayStats.bExecute S= NOT DisplayStats.bBusy AND NOT DisplayStats.bError;
DisplayStats.bExecute R= DisplayStats.bBusy OR DisplayStats.bError;

DisplayStats.sLine1 := 'PMPS-ARBITER-K';
fbFormat(sFormat := 'Fast Faults: %d', arg1:=F_ULINT(PMPS_GVL.AccumulatedFF), sOut=>DisplayStats.sLine2, bError => bError, nErrID => nErrID );

DisplayStats(eMode:=E_CX2100_DisplayModesWr.eCX2100_WriteLines);
*)

END_PROGRAM

// ---- POUs/FB_BeamClassOutputs.TcPOU
(*
Sets the beam class assertion lines for a given beam class.
*)
FUNCTION_BLOCK FB_BeamClassOutputs
VAR_INPUT
    BP : ST_BeamParams;
END_VAR
VAR_OUTPUT
END_VAR
VAR
    nBeamClass   :    BYTE;
    wBeamClass    :    BYTE;

    InitCounter: BYTE;
    counter    :    INT;

    // Beam class lines are restricted to 8 channels in the current design, since
    // there are no plans to use all 16. Channels 1-7 may be allocated to any other
    // beam classes so long as they are ordered least to greatest.
    // Channel 8 is reserved for full beam.
    {attribute 'pytmc' := 'pv: BeamClassChannel
        io: i
        field: DESC Hardwire channel state'}
        epicsBitmap : WORD;

    {attribute 'TcLinkTo' := '[1] := TIIB[PMPS_Premp]^Channel 1^Output;
                              [2] := TIIB[PMPS_Premp]^Channel 2^Output;
                              [3] := TIIB[PMPS_Premp]^Channel 3^Output;
                              [4] := TIIB[PMPS_Premp]^Channel 4^Output;

                              [5] := TIIB[PMPS_Premp]^Channel 5^Output;
                              [6] := TIIB[PMPS_Premp]^Channel 6^Output;
                              [7] := TIIB[PMPS_Premp]^Channel 7^Output;
                              '} // 8 - Full beam
    q_BC_ASSERTION_LINES    AT    %Q*    : ARRAY [1..MAX_BEAM_CLASS_LINES] OF    BOOL;
END_VAR
VAR CONSTANT
    MAX_BEAM_CLASS_LINES : BYTE := 8;
    BC_1HZ : BYTE := 1;
    BC_10HZ : BYTE := 2;
    BC_FULL : BYTE := 16;
END_VAR


// Determine BC
IF BP.nRate >= 120 THEN
    nBeamClass := BC_FULL;
ELSIF BP.nRate >= 10 THEN
    nBeamClass := BC_10HZ;
ELSIF BP.nRate >= 1 THEN
    nBeamClass := BC_1HZ;
ELSE
    nBeamClass := 0;
END_IF


//Assert Beam Class
////////////////////////////////////
//0x0 = 0000 0000 0000 0000
//0x1 = 0000 0000 0000 0001
//0xF = 1111 1111 1111 1111

//Initialize BC lines to zero on every pass
FOR InitCounter := 1 TO MAX_BEAM_CLASS_LINES DO
    q_BC_ASSERTION_LINES[InitCounter] := FALSE;
END_FOR

//Set BC lines according to beam class
//A BC of 0x0 would pass over this loop, setting none of the lines high
// , as FOR loops check the initialized variable at the top to see if it's >
// than the "TO" variable.
FOR wBeamClass:=1 TO MIN(MAX_BEAM_CLASS_LINES-1, nBeamClass) DO
    q_BC_ASSERTION_LINES[wBeamClass] := TRUE;
END_FOR

q_BC_ASSERTION_LINES[8] := nBeamClass = 16; //Set channel 8 true if BC is 16


// Readbacks for EPICS
epicsBitmap.0 := q_BC_ASSERTION_LINES[1];
epicsBitmap.1 := q_BC_ASSERTION_LINES[2];
epicsBitmap.2 := q_BC_ASSERTION_LINES[3];
epicsBitmap.3 := q_BC_ASSERTION_LINES[4];

epicsBitmap.4 := q_BC_ASSERTION_LINES[5];
epicsBitmap.5 := q_BC_ASSERTION_LINES[6];
epicsBitmap.6 := q_BC_ASSERTION_LINES[7];
epicsBitmap.7 := q_BC_ASSERTION_LINES[8];

END_FUNCTION_BLOCK
